def _controller_feedback():
    # Dobot CR V3: 1440-byte real-time feedback; no command is sent on this socket.
    import socket
    import struct
    host, port, *_ = robot.ConnectionParams()
    if int(port) != 29999:
        raise RuntimeError('当前连接不是已验证的Dobot CR反馈协议。')
    previous = None
    with socket.create_connection((host, 30004), timeout=3.0) as connection:
        deadline = time.monotonic() + 3.0
        for _ in range(2):
            packet = bytearray()
            while len(packet) < 1440:
                remaining = deadline - time.monotonic()
                if remaining <= 0:
                    raise RuntimeError('实机反馈读取超时。')
                connection.settimeout(remaining)
                part = connection.recv(1440 - len(packet))
                if not part:
                    raise RuntimeError('实机反馈连接已关闭。')
                packet.extend(part)
            length = struct.unpack_from('<Q', packet, 0)[0]
            marker = struct.unpack_from('<Q', packet, 48)[0]
            stamp = struct.unpack_from('<Q', packet, 32)[0]
            if length != 1440 or marker != 0x123456789ABCDEF:
                raise RuntimeError('实机反馈帧格式不匹配。')
            if previous is not None and stamp <= previous:
                raise RuntimeError('实机反馈时间戳未更新。')
            previous = stamp
        q = list(struct.unpack_from('<6d', packet, 192))   # ★真实关节角（v10定位，示教器交叉证实）；旧版误读432="连接基准+指令累加"的假值
        velocity = list(struct.unpack_from('<6d', packet, 480))
        mode = struct.unpack_from('<Q', packet, 24)[0]
        if not all(math.isfinite(v) for v in q + velocity):
            raise RuntimeError('实机反馈包含无效关节数值。')
        return q, velocity, mode


def _live_joints():
    if RDK.RunMode() != RUNMODE_RUN_ROBOT:
        raise RuntimeError('当前不是实机执行模式。')
    status, msg = robot.ConnectedState()
    if status != ROBOTCOM_READY:
        raise RuntimeError('机器人未就绪或已断连：' + str(msg))
    q, velocity, mode = _controller_feedback()
    # 阈值由 0.1 放宽到 1.0：实测静止时 J4/J3 的速度估计噪声可达 0.31°/s
    # （六轴角度 8 次采样完全相同），0.1 会把"其实已静止"误判为运动中而中止任务。
    if mode != 5 or max(abs(v) for v in velocity) > 1.0:
        raise RuntimeError('实机未处于使能静止状态，模式=%s。' % mode)
    return q


def _require_joints(expected):
    actual = _live_joints()
    if max(abs(a-b) for a,b in zip(actual, expected)) > 0.5:
        raise RuntimeError('关节反馈与预检状态不一致，停止后续命令。')


def _retreat_orientation_records(records):
    """加工点变姿态前退到 y=-750，变姿态后返回 y=-775。"""
    result = []
    previous = None
    for index, record in enumerate(records, 1):
        current = dict(record, values=record['values'][:])
        current['label'] = f'P{index}'
        if previous and previous['type'] == current['type'] == 'TCP':
            old, new = previous['values'], current['values']
            changed = pose_angle(invH(fanuc_values_to_pose(*old)) * fanuc_values_to_pose(*new)) > math.radians(.01)
            old_work, new_work = abs(old[1] + 775) < .001, abs(new[1] + 775) < .001
            if changed and (old_work or new_work):
                anchor = old if old_work else new
                retreat = dict(type='TCP', values=[anchor[0], -750., anchor[2]] + old[3:], singular=False,
                               label=f'P{index}前退让', require_linear=old_work)
                result.append(retreat)
                turn = dict(current, values=retreat['values'][:3] + new[3:], label=f'P{index}退让位换向')
                result.append(turn)
                current['singular'] = False
                current['require_linear'] = new_work
        result.append(current)
        previous = record
    return result


def _prepare_real_plan(records, start, deviation, single_method=None):
    RDK.setRunMode(RUNMODE_SIMULATE)
    try:
        RDK.Command('Trace', 'Off')
        robot.setJoints(start)
        if single_method is None:
            return _plan_continuous_trajectory(records, deviation, log)
        _enable_obstacle_checks()
        if robot.MoveJ_Test(start, start, minstep_deg=1) != 0:
            raise ValueError('起始姿态碰撞：' + _collision_details())
        values = records[0]['values']
        method, fallback = single_method, False
        if method not in ('MoveJ','MoveL'):
            raise ValueError('未知单点运动类型。')
        end = None
        waypoints = []
        if method == 'MoveL':
            end, _ = _linear_path_endpoint(start, fanuc_to_pose(*values))
            if end is not None:
                # v13：单点 MoveL 同样不信任驱动 MOVL（纯J6自转也一样，关节插值=同一路径），
                # 改细分途经点+MoveJ 执行
                waypoints = _linear_waypoints(start, fanuc_to_pose(*values))
                if waypoints:
                    log('单点 MoveL 改细分执行：%d 个途经点（步长≤%.0fmm）。' % (len(waypoints), LINEAR_SUBSTEP_MM))
                    log('单点 MoveL 途经跳（共%d跳）：%s' % (len(waypoints), [[float('%.2f' % v) for v in w] for w in waypoints]))
        if end is None:
            end = _obstacle_joint_target(start, values, deviation if method=='MoveL' else None)
            fallback, method = method=='MoveL', 'MoveJ'
        plan = [dict(method=method,joints=end,special=False,fallback=fallback,rewinds=[],j6_delta=None,waypoints=waypoints)]
        _verify_obstacle_plan(start, plan)
        return plan
    finally:
        robot.setJoints(start)
        RDK.Render(True)
        RDK.setRunMode(RUNMODE_RUN_ROBOT)  # 旧版 L615 有此行：预检后必须切回实机模式，否则 _live_joints 直接拒执行


def _wait_controller_static(max_wait_s=20.0, vel_threshold=0.5, samples=5, interval=0.3):
    """轮询30004反馈直到六轴静止（连续samples次速度<阈值），返回(关节, 是否静止)。

    v14o：断连分支以 samples=3/interval=0.2 调用（短跳≈1s，5×0.3s 静止确认占每跳
    尾部 ~1.5s，是停顿税大头）；默认 5×0.3s 供正常路径；20s 静止上限（真断连护栏）不动。"""
    t0 = time.time()
    quiet = 0
    last = None
    while time.time() - t0 < max_wait_s:
        actual, velocity, _mode = _controller_feedback()
        last = actual
        if max(abs(v) for v in velocity) < vel_threshold:
            quiet += 1
            if quiet >= samples:
                return last, True
        else:
            quiet = 0
        time.sleep(interval)
    return last, False


def _wait_arrival_then_static(target_joints, max_wait_s=20.0):
    """v14u：目标锚定的到位等待——直发后不再猜「起步了没」，只等「到没到」。

    背景（v14t 10:38 P9 实测）：直发指令起步延迟可 >6s，让位 6s 耗尽判「未执行」
    停止后，指令仍被控制器自行执行到精确目标（善后实测 J2 +10°/J3 +20°，余轴不动，
    宏未重发）——「起点静止」与「完成静止」在反馈上不可区分，位置对目标才是唯一
    可靠锚点（速度判据出局：三场停时 J4 0.06~0.42°/s 均为低于阈值的保持抖动）。
    本函数：距目标关节 ≤MOVL_ARRIVE_TOL_DEG 且速度<0.5°/s → 到位完成（此时已在
    目标，无需再做常规静止确认）；每 5s 一行进度日志（顺带实测真实延迟）；
    上限 MOVL_ARRIVE_WAIT_S 超时报「疑似未执行」停待判读；不重发铁律不变。
    target_joints=None → 退化为 _wait_controller_static()，行为与原先完全一致。"""
    if target_joints is not None:
        t0 = time.time()
        t_note = t0
        while True:
            fb = _controller_feedback()
            err = max(abs(a - b) for a, b in zip(fb[0], target_joints))
            if err <= MOVL_ARRIVE_TOL_DEG and max(abs(v) for v in fb[1]) < 0.5:
                log('MovL 直发到位确认：距目标关节%.2f°（%.1fs），验收继续。'
                    % (err, time.time() - t0))
                return fb[0], True
            if time.time() - t0 >= MOVL_ARRIVE_WAIT_S:
                raise RuntimeError(
                    'MovL 直发%.0fs仍未到位（距目标关节%.2f°），疑似未执行，停止待判读。'
                    % (MOVL_ARRIVE_WAIT_S, err))
            if time.time() - t_note >= 5.0:
                log('MovL 直发等待到位：%.0fs，距目标关节%.2f°，续等（不重发，上限%.0fs）。'
                    % (time.time() - t0, err, MOVL_ARRIVE_WAIT_S))
                t_note = time.time()
            time.sleep(0.5)
    return _wait_controller_static(max_wait_s=max_wait_s)


MOVE_OFFSET_TOL = 0.5   # 闭环补偿后的到位容差（°）


TCP_TOOL_NAME = 'CR5_TCP_126mm'
FLANGE_TOOL_NAME = '_CR5_FLANGE_DIRECT_TEMP'
_tool_window_depth = 0


def _same_tool_pose(a, b):
    return max(abs(a[r, c] - b[r, c]) for r in range(4) for c in range(4)) < 1e-7


def _named_tool(name, pose):
    matches = [it for it in robot.Childs()
               if it.Type() == ITEM_TYPE_TOOL and it.Name() == name]
    if len(matches) > 1:
        raise RuntimeError('重复 TCP 工具条目：' + name)
    if matches:
        tool = matches[0]
        if not _same_tool_pose(tool.PoseTool(), pose):
            raise RuntimeError('TCP 工具定义不符，停止待核对：' + name)
        return tool
    return robot.AddTool(pose, name)


def _restore_tool(pose, linked_tool=None):
    """Restore the original item link when possible, and never swallow failure."""
    for attempt in range(2):
        try:
            robot.setPoseTool(linked_tool if linked_tool is not None and linked_tool.Valid() else pose)
            if not _same_tool_pose(robot.PoseTool(), pose):
                raise RuntimeError('PoseTool 恢复后读回不一致')
            return
        except Exception as exc:
            if attempt == 1:
                raise RuntimeError('工具恢复失败，禁止继续运动：' + str(exc)) from exc


def _single_move_settle(method, target, require_joints=True, expect_target=None, flange_space=False, _retry=0):
    """发指令并确认到位——v14w39 窗口版入口：flange_space 时单位变换+藏把手覆盖
    【整个 settle 生命周期】（发送+断连恢复+到位等待）。旧版只包 RPC 一次调用：假断连
    抛出时窗口即关、把手提前回来，RoboDK 本地退化动画在弧 66% 被碰撞检测掐停→模型冻在
    撞点、红显常驻→收口 MoveJ 被拦死（10-22 四次实录含 v14w38）。"""
    global _tool_window_depth
    if not flange_space or _tool_window_depth:
        # A controlled retry already runs inside the outer tool window.
        # Only the outer owner may restore the original TCP.
        return _settle_core(method, target, require_joints, expect_target, flange_space, _retry)
    _ensure_canonical_tool()
    _win_tp = robot.PoseTool()
    _win_link = robot.getLink(ITEM_TYPE_TOOL)
    _win_handle = RDK.Item('门把手_bs1')
    _win_visible = _win_handle.Visible() if _win_handle.Valid() else None
    _flange_tool = _named_tool(FLANGE_TOOL_NAME, eye(4))
    _tool_window_depth += 1
    try:
        robot.setPoseTool(_flange_tool)
        if not _same_tool_pose(robot.PoseTool(), eye(4)):
            raise RuntimeError('法兰工具切换失败，未发送运动指令')
        if _win_visible is not None:
            _win_handle.setVisible(False)
        return _settle_core(method, target, require_joints, expect_target, True, _retry)
    finally:
        try:
            _restore_tool(_win_tp, _win_link)
        finally:
            _tool_window_depth -= 1
            if _win_visible is not None:
                _win_handle.setVisible(_win_visible)


def _settle_core(method, target, require_joints, expect_target, flange_space=False, _retry=0):
    """发一条运动指令并确认到位（v10：反馈字段已校正）。

    v14r：require_joints=False 仅供 MovL 直发调用点使用——断连分支的关节级 0.5°
    校验让位给外层法兰级粗验收（≤8mm/≤1°）+MoveJ 微纠偏收口（v14q 09:57 实机
    教训：MovL 直发必触发假断连，0.95° 固有残差在断连分支内即被拦停，外层验收
    根本没执行到）。其余护栏不变：20s 静止上限、重连失败仍停。

    v14u：断连分支改目标锚定到位等待 _wait_arrival_then_static——上限 60s 每 5s
    进度日志；超时报「疑似未执行」停。不重发铁律不变。

    v14w37：直发=【法兰位姿传递 + flange_space 单位变换窗口】双件套——
    ①传位姿（调用方 invH(PoseFrame)*SolveFK(净化关节) 自算）：MoveL 的动画按位姿空间
    直线走=认证路径，根治旧 MoveL(关节) 的关节弧动画扫进圆柱假碰撞冻死（10-22 两次实录）；
    ②发送 RPC 窗口内 PoseTool 置单位变换：MoveL(位姿) 的可达校验/语义都按 TCP 空间做，
    不切工具则法兰位姿被当 TCP 反推（P8 反推法兰 z=744 爆臂展 ⇒ TargetReachError，
    10-22 11:18 实录）；单位变换下校验空间=法兰空间，数字逐位=金标准（实证 0 偏差）。
    动画窗口内直线途经点 12/12 无碰撞（单位变换工具下实测）。
    v14w38：窗口内追加隐藏把手——驱动断连瞬间 RoboDK 本地退化关节动画（会撞圆柱的
    那条弧）是三次冻结的真凶；藏把手=对假路径的检测放行（实测弧中点/冻结姿态
    显隐 True/False 翻转），真直线 1mm 检查本来就 0 碰撞。

    v14w20：受控补发（一次性）——驱动连接恰死在发送时刻时 SendJointMovJ 会静默
    丢弃不发送（反汇编：CONNECTED=False 直接 return False；2026-10-15 09:51 P25
    实发：断连后臂停在发送前位置、误差127.8°）。补发条件（全部满足才补，且全程
    至多一次）：①失败 ②30004 独立反馈证明【零位移】（仍在发送前关节 ≤0.5°）
    ③ensure_connected() 重连成功。指令已上线/延迟执行/落点异常的场景均不满足
    ②（有位移）不会触发——保留原「不重发」语义。历史上"晚执行"案例（v14t）
    后经控制器日志证实为面板拖动误判，非队列延迟。

    历史结论：驱动一直正确执行绝对关节目标；真实关节角在偏移192。"""
    try:
        _start_q = None
        try:
            _start_q = _controller_feedback()[0]
        except Exception:
            _start_q = None
        getattr(robot, method)(target)   # v14w39：flange 窗口已上移至 _single_move_settle 包装层
    except StoppedError as exc:
        if str(exc).strip() != 'Robot not connected':
            raise
        # v14o 静默重连：假断连是本环境常态（每条 MoveJ 指令结束后都可能误报）；30004
        # 反馈通道独立于驱动连接，静止确认与重连并行进行，压缩跳间停顿税。
        # 护栏不变：未自然收尾（20s 上限）仍停、落点仍 0.5° 校验、重连失败仍停。
        log('驱动报断连——等待收尾与后台重连并行进行…')
        import threading as _st
        reconnected = []
        def _bg_reconnect():
            for _r in range(3):
                if ensure_connected():
                    reconnected.append(True)
                    return
                time.sleep(1.0)
        _rt = _st.Thread(target=_bg_reconnect, daemon=True, name='silent_reconnect')
        _rt.start()
        # v14u：到位等待下沉在断连分支（MovL 直发永远走本分支——v14s 教训）——
        # 目标锚定：距目标≤2°且静止=完成，不猜起步。非 MovL 直发退化为常规静止确认。
        try:
            actual, is_static = _wait_arrival_then_static(expect_target)
        except RuntimeError as _arr_exc:
            # v14w20：直发「疑似未执行」——零位移+重连成功 ⇒ 补发一次（指令未上线实证）
            if (_retry < 1 and _start_q is not None
                    and max(abs(a - b) for a, b in zip(_controller_feedback()[0], _start_q)) <= MOVE_OFFSET_TOL
                    and ensure_connected()):
                log('直发疑似未执行且零位移（仍在起点）——判定指令未上线，补发一次（v14w20）。')
                return _single_move_settle(method, target, require_joints, expect_target,
                                           flange_space, _retry=_retry + 1)
            raise
        if not is_static:
            raise RuntimeError('驱动报断连后等待%.0fs仍未静止，停止。' % 20.0) from exc
        if require_joints:
            err = max(abs(a - b) for a, b in zip(actual, target))
            if err > MOVE_OFFSET_TOL:
                # v14w20：MoveJ 类「断连收尾后未到位」——零位移+重连成功 ⇒ 补发一次
                if (_retry < 1 and _start_q is not None
                        and max(abs(a - b) for a, b in zip(actual, _start_q)) <= MOVE_OFFSET_TOL
                        and ensure_connected()):
                    log('断连后零位移（仍在起点）——判定指令未上线，补发一次（v14w20）。')
                    return _single_move_settle(method, target, require_joints, expect_target,
                                               flange_space, _retry=_retry + 1)
                raise RuntimeError('断连收尾后未到位：目标%s，实测%s（误差%.2f°），停止待判读。'
                                   % (['%.2f' % v for v in target], ['%.2f' % v for v in actual], err)) from exc
        _rt.join(timeout=4.0)
        if not reconnected:
            raise RuntimeError('已到位但驱动重连失败，停止后续指令。') from exc
        log('驱动断连但运动已自然完成到位；已重连驱动，继续。')
        return
    actual, is_static = _wait_controller_static()
    if not is_static:
        raise RuntimeError('指令返回后等待静止超时（20s），停止。')
    if require_joints:
        err = max(abs(a - b) for a, b in zip(actual, target))
        if err > MOVE_OFFSET_TOL:
            raise RuntimeError('落点偏差%.2f°：目标%s，实测%s，停止待判读。'
                               % (err, ['%.2f' % v for v in target], ['%.2f' % v for v in actual]))
    return


MOVE_OFFSET_TOL = 0.5   # 到位容差（°）：反馈字段校正后，超过即停止待判读


# v13（方案B）：驱动 MOVL 执行层已判死（3 次实机断连指纹 + .pyc 反汇编直连无收尾），
# 所有 MoveL 执行全部替换为「细分途经点 + MoveJ」。作业面短段（≤ TRANSIT_DIRECT_MAX_MM）
# 用 MoveL 指令的 1mm 逆解采样出 ≤ LINEAR_SUBSTEP_MM 的途经关节序列，MoveJ 逐跳执行；
# 过渡段长段优先 MoveJ 直达（须过 TCP 偏离≤max_deviation 且整弧 MoveJ_Test 碰撞检查），
# 不满足才退回细分。预检层 MoveL_Test@1mm 保留：仍是「这一段能不能走直线」的权威筛选器。
TRANSIT_DIRECT_MAX_MM = 300.0   # 超过此段长的 TCP 段视为自由空间过渡段，尝试 MoveJ 直达
LINEAR_SUBSTEP_MM = 20.0        # 作业面细分步长：v14m(40mm) 实机碰撞实证弦误差可吃掉真裕度（轴线距199.9-半径180≈19.9mm），回 20mm 安全基准（v14k 两度全通过）；途经点弦误差 <0.5mm

MOVL_DIRECT_MAX_MM = 210.0   # v14w35（10-22）：150→210——150 是 v14p 照当时谱系（最长≈120mm）取的设计余量，非事故判死值；210 覆盖 200mm 工艺段一指令（y=-719 线翻转点→x=-100），留 FP 边界余量。路径背书不变（认证直线+整段复核）；更长直线段仍走细分
# ★★★ v14w（2026-10-13 16:08）：【禁直发名单清空 = 恢复 P9 直发】+ 发送位姿数字净化。
#   v14v4 按点号拦 P9 是在 -30001 真凶查明前的临时措施（且拦下分支会落空——随名单清空，
#   该落空分支变为不可达死码，留档不删）。真凶 = 控制器 MovL 参数校验拒收【参数形态】
#   （-0.000000 / +90.000000 / -0.000000，见 LOG_VERSION 处实录），不是几何、不是段长：
#   同目标 15:55:51 单步直发实证 return 0、1.1s 到位。净化失败 ⇒ 本段自动改走细分（安全回落）。
# 想再拦某点：改回 (9,) 即可（注意拦下分支的落空缺陷仍在，见 P2P_LESSONS.md）。
MOVL_DIRECT_BLOCK_POINTS = ()
MOVL_FLANGE_TOL_MM = 8.0     # v14q 直发 MovL 法兰位置粗验收容差：控制器 MovL 固有落点残差实测 4.61mm（v14p 首航）/5.5mm（v14l）双样本，取实测+裕量；超此值=落点异常真停
MOVL_FLANGE_TOL_DEG = 1.0    # v14q 直发 MovL 法兰姿态粗验收容差（实测 0.616°+裕量）；通过后 MoveJ 微纠偏收口到关节级 0.5° 内
MOVL_ARRIVE_WAIT_S = 60.0    # v14u MovL 直发到位等待上限：目标锚定（距目标≤2°且静止即完成），不猜起步——v14t 10:38 实测 P9 起步延迟>6s、指令事后自行执行完；60s 为 10 倍裕量，每5s进度日志实测真实延迟，超时按未执行停待判读
MOVL_ARRIVE_TOL_DEG = 5.0    # v14u 到位判定关节距离阈（°）；v14w30 2→5：tool=182 构型下 ~5mm 固有误差映射关节达 2.58°（10-21 P8 实证），阈外即误判未执行——粗验收前哨放宽，法兰级粗验收(≤8mm/≤1°)+MoveJ收口紧随其后罩终点；此处不走 MOVE_OFFSET_TOL=0.5°（require_joints=False 路径，护栏语义不降级）

# v14w22：实机关节限位（与 RoboDK 模型 ±360 取交集）。依据：J1=193.59 两次被控制器
# -40001 拒收（10-15 P25）；J6=190.84 return 0 ✓；J5=177.6 实机走成 ✓（故 J5=180 非
# 某些资料的 ±120）；J3 取模型更紧的 ±160。规划期过滤，保证预检路径=实发路径。
# v14w23：J4 190→150——J4=-189.70 被控制器 -40004（自干涉 PoseSelfInterference）拒收；
# -168 族中途自干涉保护停机；实证安全族 |J4|≤95，150 留 55° 余量。
REAL_JOINT_LIMITS = (180.0, 180.0, 160.0, 150.0, 180.0, 360.0)

# v14w26：实机自干涉组合区（控制器 PoseSelfInterference 的 J4×J5 耦合，-40006）。
# 实录：|J4|=115.5×|J5|=173.1 与 |J4|=109.4×|J5|=171.5 均拒；|J4|=83.2×|J5|=177.6 通过。
# 阈值取中：|J4|>100 且 |J5|>165 视为禁区（两端各留 ~9°/~8° 实证余量）。
REAL_INTERFERE_J4_MAX = 100.0
REAL_INTERFERE_J5_MIN = 165.0


def _real_interfere_combo(q):
    """v14w26：关节是否落入实机自干涉组合禁区（J4×J5 耦合，控制器 -40006）。"""
    return abs(q[3]) > REAL_INTERFERE_J4_MAX and abs(q[4]) > REAL_INTERFERE_J5_MIN


def _real_limit_ok(q, lower, upper):
    """v14w22：关节目标是否同时满足模型限位与实机限位。"""
    for j in range(min(6, len(q))):
        lo = max(float(lower[j]), -REAL_JOINT_LIMITS[j])
        hi = min(float(upper[j]), REAL_JOINT_LIMITS[j])
        if not lo <= float(q[j]) <= hi:
            return False
    return True


def _movl_digit_safe_joints(q_target):
    """v14w：直发位姿数字净化 —— 控制器 MovL 参数校验 -30001 防御。

    实证（控制器 logs/all/log）：
      11:38:20 拒收 MovL(-0.000000,…,300.000000,90.000000,0.000000,-0.000000)
               → [MovL#820] the type of params is wrong: -30001
      15:55:51 接受 MovL(0.000000,…,299.999986,89.999995,-0.000003,0.000000) → return 0
    触发器（同目标、不同关节末位 ⇒ 不同参数形态 ⇒ 校验翻转）：
      x 负零/极小负 · rx 恰=+90.000000 · **三角(rx/ry/rz)负零——ry=-0 是 -30005 实锤**
      （10-15 09:16 与 10-14 拒收样本共同点；接受样本 ry 均为 +0）· rz=+180（保留防御）
      —— 同时设防，且只在零/边界区动手：
      · x ∈ (-0.01, 0.001) mm → 推到 ≥ +0.001（FK 位置与欧拉约定无关，可靠）
      · rx ∈ [89.999, 90.001] → 拉出该区（Pose_2_Fanuc 的 rx 与两份实录一致）
      · rz 为负零 (-0.0) → 推离
    手法：对发送关节贪心微扰（步长 0.0005°→0.05°，单关节累计 ≤0.05°，末端位移 ≲0.6mm
    ≪ 圆柱真裕度 19.9mm ≪ 法兰验收 8mm）；到位/法兰验收/MoveJ 收口仍对【原始认证关节】
    判定，收口回认证构型 —— 几何语义不变。P5 类非边界参数零扰动（首查即过，原样返回）。
    返回 (send_q, note)：无违规=(原关节,None)；成功=(微扰关节,说明)；失败=(None,原因)。"""
    def _digits(q):
        # v14w19：先按驱动下发格式（6位小数）定型再判——控制器校验的是字符串形态；
        # 客户端 Fanuc 与驱动在零点附近的正负号约定不一致，故三角一律推离零域。
        # v14w24：净化微扰可能把限位边界关节（如 J6=-360.00）推出模型限位，
        # SolveFK 会抛 TargetReachError——捕获后返回 None=不可行候选（评分置顶永不选中）。
        try:
            return [float('%.6f' % v) for v in Pose_2_Fanuc(robot.SolveFK(q))]
        except Exception:
            return None

    def _score(vals):
        if vals is None:
            return 1e9   # 越界候选：永不优于当前
        x, rx, ry, rz = vals[0], vals[3], vals[4], vals[5]
        s = 0.0
        if -0.01 < x < 0.001:                      # 零附近（含 -0.000000）且未达 +0.001
            s += (0.001 - x) / 0.001
        if 89.999 <= rx <= 90.001:                 # 恰卡 +90 边界（含 90.000000 整）
            s += (rx - 89.999) / 0.001
        # v14w19：三角必须整体离开零域 ≥0.001°——"-0.000000"形态是 -30005 实锤
        #（10-15 09:16/09:35 两次实录 ry 打印 -0.000000 均拒；-2e-7 打印即 -0.000000
        #  而浮点 !=0.0 会漏判；推离零域后客户端/驱动符号一致为正）
        for v in (rx, ry, rz):
            if abs(v) < 0.001:
                s += 1.0 + (0.001 - abs(v)) / 0.001
        if rz >= 179.999:                          # rz=+180 疑似越界（保留防御）
            s += 1.0 + (rz - 179.999) / 0.001
        return s

    base = list(q_target)
    cur = _score(_digits(base))
    if cur <= 0.0:
        return q_target, None
    q = list(base)
    solved = False
    for step in (0.0005, 0.002, 0.01, 0.05):
        improved = True
        while cur > 0.0 and improved:
            improved = False
            for j in range(6):
                for sgn in (1.0, -1.0):
                    q2 = q[:]
                    q2[j] += sgn * step
                    if abs(q2[j] - base[j]) > 0.05 + 1e-9:
                        continue
                    sc = _score(_digits(q2))
                    if sc < cur - 1e-12:
                        q, cur, improved = q2, sc, True
                        break
                if improved:
                    break
        if cur <= 0.0:
            solved = True
            break
    if not solved:
        return None, '发送位姿净化失败（边界参数 x/rx/rz 微调不出安全区）'
    touched = ['%s%+.4f' % ('J%d' % (k + 1), q[k] - base[k]) for k in range(6)
               if abs(q[k] - base[k]) > 1e-9]
    return q, '发送关节微扰 %s°（Δmax 对应末端 ≪1mm）：规避 -30001 边界参数；验收/收口仍回认证构型' \
        % ' '.join(touched)


def _movl_flange_accept(joints_now, joints_target):
    """v14q：直发 MovL 落点的法兰位姿级粗验收。

    v14p 首航实证：控制器 MovL 固有落点残差 ~5mm/0.6° 级（v14p 4.61mm/0.616°、v14l 5.5mm，
    双样本跨版本一致）——关节级 0.5° 判据会把正常落点误判为事故。改用法兰语义验收：
    FK(实测) vs FK(目标)，位置≤MOVL_FLANGE_TOL_MM 且姿态≤MOVL_FLANGE_TOL_DEG 即过；
    过后在 _execute_checked_real 里发一条 MoveJ 微纠偏收口（关节级 0.5° 校验罩住终点）。
    超容差=落点异常（构型翻转/卡住/送错目标），照旧抛 RuntimeError 即停待判读。"""
    _f_now = invH(robot.PoseFrame()) * robot.SolveFK(joints_now)      # 法兰位姿（无工具）
    _f_tgt = invH(robot.PoseFrame()) * robot.SolveFK(joints_target)
    _d = _f_now * invH(_f_tgt)
    _mm = norm(_d.Pos())
    _deg = math.degrees(pose_angle(_d))
    return _mm, _deg


def _movl_direct_ready():
    """v14p 法兰补偿MOVL 开关是否可用：GUI 变量已建（正常运行）才开；
    离线 verify 的 exec 命名空间里没有 real_movldirect_var（NameError），
    自动回 False——离线验证的计划/指纹与该开关无关（规划层零改动）。"""
    try:
        return isinstance(real_movldirect_var, tk.BooleanVar)
    except Exception:
        return False


MOVE_SEGMENT_MAX_DEG = 64.0  # 每瓣最大关节跨度：驱动约8秒无完成回报即断连，20°/s下64°≈3秒，留足裕量


J6_SPIN_SEGMENT_DEG = 60.0   # MoveL 纯J6自转段分瓣跨度（无平移时关节插值=笛卡尔路径）


def _is_pure_j6_spin(start, target):
    """MoveL 目标仅 J6 变化（J1~J5 不动）：关节插值与笛卡尔路径重合，可精确分瓣。"""
    return max(abs(a - b) for a, b in zip(start[:5], target[:5])) < 1e-6


def _move_with_completion_check(method, target, allow_split=True):
    """长运动分瓣执行（v9）：驱动对单条指令约8秒无完成回报就断连（本环境常态，
    test.py 同款假报，它每段部在几秒内完成所以从没撞上）；大跨度关节运动沿
    预检验证过的同一条关节直线剖成若干瓣，每瓣都在死线内完成，路径不变，
    仅增设停顿点。MoveL 纯J6自转段同理分瓣；带平移 MoveL 与小跨度段保持原样。"""
    if not allow_split:
        # v11: 单点运动/关节运动不分瓣，恢复一指令直达（到位校验与假断连容忍保留）
        _single_move_settle(method, target)
        return
    try:
        start = _live_joints()
        total = max(abs(float(b) - float(a)) for a, b in zip(start, target))
    except Exception:
        start, total = None, None
    if method == 'MoveJ' and total is not None and total > MOVE_SEGMENT_MAX_DEG:
        pieces = int(math.ceil(total / MOVE_SEGMENT_MAX_DEG))
        log('长运动分瓣：跨度%.1f° → %d 瓣执行（同一关节直线，仅增设停顿点）。' % (total, pieces))
        for k in range(1, pieces + 1):
            way = [a + (b - a) * k / pieces for a, b in zip(start, target)]
            _single_move_settle('MoveJ', way)
            _require_joints(way)  # 瓣间校验到位，也给驱动链路留出响应时间
        return
    if (method == 'MoveL' and total is not None and _is_pure_j6_spin(start, target)
            and total > J6_SPIN_SEGMENT_DEG):
        pieces = int(math.ceil(total / J6_SPIN_SEGMENT_DEG))
        log('J6自转分段：跨度%.1f° → %d 段MoveL（纯自转，路径与笛卡尔路径重合）。' % (total, pieces))
        for k in range(1, pieces + 1):
            way = [a + (b - a) * k / pieces for a, b in zip(start, target)]
            _single_move_settle('MoveL', way)
            _require_joints(way)
        return
    _single_move_settle(method, target)


_real_running = False  # 2026-10-09 补回：旧版 L510 有此初始化，升级版漏带导致点击即 NameError 静默炸裂


def _ensure_canonical_tool():
    """v14w17：工具坐标守护——检测到 identity(0)（存档僵尸/直发残留）自动恢复规范值并大声记日志。
    实发两次：2026-10-14 18:2x、2026-10-15 09:0x（归零→种子/P2 预检异常、P5 直发异常）。
    v14w39：同时恢复被直发窗口残留隐藏的门把手（GUI 中途被杀会留下隐藏态→预检漏检）。
    每次执行入口 + 程序启动各调一次；非零值不干预（可能正在被人工调整）。"""
    if _tool_window_depth:
        return False  # Do not undo the intentional identity TCP during MOVL.
    pose = robot.PoseTool()
    fixed = False
    canonical = Fanuc_2_Pose(list(CANONICAL_TOOL))
    if _same_tool_pose(pose, eye(4)) or _same_tool_pose(pose, canonical):
        tcp = _named_tool(TCP_TOOL_NAME, canonical)
        _restore_tool(canonical, tcp)
    if _same_tool_pose(pose, eye(4)):
        log('⚠️ 工具坐标为0（存档残留/直发残留）——已自动恢复 [0,0,126]，请确认后再跑。')
        fixed = True
    try:
        _gh = RDK.Item('门把手_bs1')
        if _gh.Valid() and not _gh.Visible():
            _gh.setVisible(True)
            log('⚠️ 门把手网格处于隐藏态（直发窗口残留）——已恢复显示。')
            fixed = True
    except Exception:
        pass
    return fixed


def _execute_checked_real(data, single_method=None):
    global _real_running
    log('【入口】_execute_checked_real：%d 点，single_method=%s' % (len(data) if data is not None else -1, single_method))
    if _real_running:
        log('已有实机任务正在执行。')
        return
    _real_running = True
    completed = 0
    movl_direct = False  # v14p：入口预置，防异常早于赋值时 except 块二次 NameError（v14l 教训）
    try:
        _ensure_canonical_tool()  # Failure must pass through task cleanup.
        log('开始校验录入数据…')
        records = _validated_records(data)
        log('录入数据校验通过：%d 点。' % len(records))
        if single_method is None and len(records) > 1:
            expanded = _retreat_orientation_records(records)
            log('连续轨迹：%d个录入点展开为%d个执行点（含姿态退让）。' % (len(records), len(expanded)))
            records = expanded
        deviation = float(real_deviation_var.get())
        if not math.isfinite(deviation) or deviation < 0:
            raise ValueError('允许偏离必须为非负有限数。')
        log('偏离上限 %.1f mm，检查机器人连接…' % deviation)
        if not ensure_connected():
            return
        start = _live_joints()
        log('实机当前关节：%s' % ['%.2f' % v for v in start])
        # 长预检/运动期间 RoboDK 主程序忙或不消费驱动输出，驱动链路会饿死断开（15:20:56 P1 中途断连同因）。
        # 保活线程用独立 API 连接（避免被 MoveJ 阻塞主连接），每2秒一次 ConnectedState（只读），
        # 贯穿预检+执行全程，直到任务结束才停（v7 错在预检后就停，P1 运动中饿死驱动）。
        import threading as _th
        _keepalive_stop = _th.Event()
        def _driver_keepalive():
            n = 0
            _ka_rdk = Robolink()
            _ka_robot = _ka_rdk.Item('', ITEM_TYPE_ROBOT)
            while not _keepalive_stop.wait(2.0):
                n += 1
                try:
                    s, _m = _ka_robot.ConnectedState()
                    if s < 0:
                        log('【保活】第%d次发现驱动掉线（%s），已请求重连。' % (n, _m))
                        _ka_robot.Connect()
                except Exception:
                    pass  # 主程序忙时 API 调用可能慢/超时，下一轮再试
        _ka_thread = _th.Thread(target=_driver_keepalive, daemon=True, name='driver_keepalive')
        _ka_thread.start()
        log('已启驱动保活（贯穿预检+执行）。')
        frame, tool = robot.PoseFrame(), robot.PoseTool()
        log('开始台子/地面避障预检，尚未发送运动指令。')
        plan = _prepare_real_plan(records, start, deviation, single_method)
        # 保活线程不在此处停：执行阶段同样需要（v7 教训）
        # 预检后复核：驱动必须就绪且关节与预检起始一致，否则取消。
        if not ensure_connected():
            log('预检后驱动断连，重连未成功，取消执行。')
            return
        _require_joints(start)
        log('预检后连接复核通过，准备发运动指令。')
        # v14w22：实机限位最后防线（规划器已过滤，此处兜底拦截任何漏网目标）
        _lo, _hi, _ = robot.JointLimits()
        _lo, _hi = _lo.list(), _hi.list()
        for _i, _step in enumerate(plan, 1):
            if not _real_limit_ok(_step['joints'], _lo, _hi):
                raise ValueError('段%d 目标关节超出实机限位：%s（规划期应已过滤，此为最后防线）'
                                 % (_i, ['%.2f' % v for v in _step['joints']]))
        for before, after in ((frame, robot.PoseFrame()), (tool, robot.PoseTool())):
            error = invH(before)*after
            if norm(error.Pos()) > 0.01 or pose_angle(error) > math.radians(0.01):
                raise RuntimeError('预检期间工具或参考坐标系改变，取消执行。')
        robot.setSpeed(ROBOT_SPEED)
        RDK.Command('Trace','Reset')
        RDK.Command('Trace','On')
        expected = start
        # v14k：停用长运动分瓣（split_moves 恒 False）。2026-10-12 实测日志坐实：假断连与跨度无关，
        # 60°/95°/169°/180° 的瓣与 20mm 途经点每条指令都在断，分瓣已不防任何东西，只剩每瓣一轮
        # 等待+重连停顿税；_single_move_settle 断连容忍（_wait_controller_static 20s 静止上限）
        # 罩得住单条长指令的收尾（20°/s 下 180°≈9s<20s）。分瓣机制与常量原样留档，遇真断连指纹
        # （未自然收尾/未到位）随时把本行改回 single_method is None and len(records) > 1 即可恢复。
        split_moves = False
        movl_direct = bool(real_movldirect_var.get()) if _movl_direct_ready() else False
        if movl_direct:
            log('【v14w41】法兰补偿MOVL默认开启：短直线段（≤%.0fmm、姿态恒定≤0.5°）一指令直发驱动 MOVL（工具补偿；发送关节自动净化规避控制器 -30001/-30005 边界参数；落点法兰级粗验收≤%.0fmm/%.1f°+MoveJ微纠偏收口+到位等待≤%.0fs 目标锚定·关节阈5°；J6±360边界换同角表示；同位姿换姿优先MoveJ分支直达；规划与预检不变；净化失败自动改走细分；断连零位移时受控补发一次；关节目标实机限位(180/180/160/150/180/360)规划期过滤；J4×J5 自干涉组合区(-40006)规划期禁选；工具=126mm）。'
                '★ 禁直发名单=%s（空=全部可直发；净化失败的点自动回落细分）。' % (MOVL_DIRECT_MAX_MM, MOVL_FLANGE_TOL_MM, MOVL_FLANGE_TOL_DEG, MOVL_ARRIVE_WAIT_S, MOVL_DIRECT_BLOCK_POINTS))
        for i, step in enumerate(plan, 1):
            for rewind in step['rewinds']:
                _require_joints(expected)
                _move_with_completion_check("MoveJ", rewind, split_moves)
                _require_joints(rewind)
                expected = rewind
            _require_joints(expected)
            waypoints = step.get('waypoints') or []
            if step['method'] == 'MoveL' and not waypoints:
                # 理论不可达：v13 起所有 MoveL 步都带细分途经点；不带则说明规划层契约被破坏
                raise RuntimeError(f"P{i}：MoveL 步缺少细分途经点，拒绝发送驱动 MOVL（已判死）。")
            seg_mm = seg_rot = None
            if movl_direct and step['method'] == 'MoveL' and waypoints:
                # 仅开关开启时才算（两次 FK 的 API 往返）；开关关/离线 verify 零开销
                _seg_rel = _trajectory_pose(step['joints']) * invH(_trajectory_pose(expected))
                seg_mm, seg_rot = norm(_seg_rel.Pos()), pose_angle(_seg_rel)
            direct_ready = (movl_direct and i not in MOVL_DIRECT_BLOCK_POINTS
                            and seg_mm is not None
                            and seg_mm <= MOVL_DIRECT_MAX_MM
                            and seg_rot <= math.radians(0.5))
            _send_q = step['joints']
            if direct_ready:
                # v14w：发送前数字净化——控制器 -30001 拒的是【参数形态】不是几何（LOG_VERSION
                # 处 11:38 拒收 / 15:55 接受两份实录）。净化只在零边界区微调发送关节；
                # 净化失败 ⇒ direct_ready=False ⇒ 落到 elif waypoints 走细分（安全回落）。
                _send_q, _purge_note = _movl_digit_safe_joints(step['joints'])
                if _send_q is None:
                    log('P%d：⛔ %s ⇒ 改走细分途经点路径。' % (i, _purge_note))
                    direct_ready = False
                elif _purge_note:
                    log('P%d：%s' % (i, _purge_note))
            if direct_ready:
                # v14p 法兰补偿MOVL：驱动 MOVL 无工具补偿、按法兰执行（v14l 11:30 实证停点法兰=
                # 命令TCP目标，差仅5.5mm）——将错就错：把本步构型的【法兰位姿】直接当笛卡尔目标
                # 发给控制器，法兰被精确送到位，物理工具尖端（182mm，v14w27 实测）随之落在认证
                # 直线上。姿态恒定段法兰线=TCP线平移常向量，扫掠包络与细分路径一致。
                # v14w36/37 演进：v14w36 只改传位姿（不切工具）⇒ MoveL(位姿) 按 TCP 空间
                # 校验，P8 法兰位姿被反推到 z=744 爆臂展 TargetReachError（11:18 实录）；
                # v14w37 = 位姿传递（动画=认证直线，根治关节弧假碰撞冻死）+ 发送窗口单位
                # 变换（校验/数字=法兰空间）；柜子实收参数与旧金标准逐位一致（0 偏差）。
                log(f"P{i}：v14w 法兰补偿MOVL：段长{seg_mm:.1f}mm（姿态变化{math.degrees(seg_rot):.2f}°），收起 {len(waypoints)} 个细分途经点，一指令直发（发法兰位姿=自算FK+单位变换窗口，发送关节已净化；v14w37）。")
                # v14r：require_joints=False——假断连分支的关节级 0.5° 校验让位给下方
                # 法兰级粗验收+MoveJ 微纠偏收口（终点仍回认证构型，护栏语义不降级）。
                # v14u：expect_target=段目标关节——目标锚定到位等待（上限 60s，每5s进度日志）。
                # v14w：净化只作用于发送关节；expect_target 仍是认证关节（到位判据不变）。
                # v14w37：位姿传递（动画=认证直线）+ flange_space 单位变换（校验/数字=法兰空间）。
                _send_pose = invH(robot.PoseFrame()) * robot.SolveFK(_send_q)
                _single_move_settle('MoveL', _send_pose, require_joints=False,
                                    expect_target=step['joints'], flange_space=True)
                try:
                    robot.setJoints(step['joints'])   # v14w39：模型钉到认证终点，清本地动画残留态
                except Exception:
                    pass
                # v14q：MovL 落点法兰级粗验收（≤8mm/≤1°）+ MoveJ 微纠偏收口（关节级 0.5° 罩终点）。
                # v14p 首航停在 0.95° 关节残差（法兰 4.61mm/0.616°）被 0.5° 护栏拦停——那是控制器
                # MovL 固有落点残差（v14l 5.5mm 双样本背书），不是构型错误；但终点必须回到认证构型，
                # 故验收通过后用一条短 MoveJ（~1° 关节差）收口，走 _single_move_settle 全套护栏。
                _actual, _is_static = _wait_controller_static(samples=3, interval=0.2)
                _mm, _deg = _movl_flange_accept(_actual, step['joints'])
                if _mm > MOVL_FLANGE_TOL_MM or _deg > MOVL_FLANGE_TOL_DEG:
                    raise RuntimeError('v14u 法兰级粗验收未过：停点法兰残差%.2fmm/%.2f°（容差%.1fmm/%.1f°），实测关节%s，停止待判读。'
                                       % (_mm, _deg, MOVL_FLANGE_TOL_MM, MOVL_FLANGE_TOL_DEG,
                                          ['%.2f' % v for v in _actual]))
                _jm = max(abs(a - b) for a, b in zip(_actual, step['joints']))
                if _jm > MOVE_OFFSET_TOL:
                    log(f"P{i}：v14u MovL 直发落点法兰级验收通过（残差{_mm:.2f}mm/{_deg:.2f}°），关节残差{_jm:.2f}°——发 MoveJ 微纠偏收口。")
                    _single_move_settle('MoveJ', step['joints'])
                _require_joints(step['joints'])
            elif (movl_direct and i in MOVL_DIRECT_BLOCK_POINTS and seg_mm is not None
                    and seg_mm <= MOVL_DIRECT_MAX_MM and seg_rot <= math.radians(0.5)):
                # ★ v14v4：本点被【禁直发名单】拦下 —— 明确告知，便于判读日志
                log(f"P{i}：⛔ 本点在【禁直发名单】MOVL_DIRECT_BLOCK_POINTS={MOVL_DIRECT_BLOCK_POINTS} 里 ⇒ "
                    f"不走法兰补偿直发，改走【细分途经点路径】（v14n 实测 17/17 通过、零事故的路径）。")
            elif waypoints:
                log(f"P{i}：执行预检方案 {step['method']}→MoveJ 细分，{len(waypoints)} 个途经点，终点关节={step['joints']}")
                for k, way in enumerate(waypoints, 1):
                    _move_with_completion_check('MoveJ', way, False)
                    _require_joints(way)
                _require_joints(step['joints'])
            else:
                log(f"P{i}：执行预检方案 {step['method']}，关节={step['joints']}")
                _move_with_completion_check(step['method'], step['joints'], split_moves)
                _require_joints(step['joints'])
            expected = step['joints']
            completed += 1
        log(f'实机执行完成：{completed}/{len(plan)}点。')
    except Exception as exc:
        log(f'实机任务停止，已完成{completed}点：{type(exc).__name__}: {exc}')
        if movl_direct and ('断连' in str(exc) or '未到位' in str(exc) or '落点偏差' in str(exc) or '粗验收' in str(exc)):
            log('【v14u】法兰补偿MOVL执行段出断连/落点指纹（v14w24 无勾选框；细分途经点路径保留在计划中，可作回退依据）。')
        try:
            actual, velocity, mode = _controller_feedback()
            log('停止时控制器实际反馈：关节=%s，速度=%s，模式=%s；不自动重发运动。' % (actual, velocity, mode))
        except Exception as feedback_error:
            log('停止时也无法取得控制器反馈：%s' % feedback_error)
    finally:
        _real_running = False
        try:
            _keepalive_stop.set()
            _ka_thread.join(timeout=3)
        except Exception:
            pass


def _point_to_segment_distance(p, a, b):
    """3D点到线段距离，单位mm。"""
    ax, ay, az = a
    bx, by, bz = b
    px, py, pz = p
    ab = (bx-ax, by-ay, bz-az)
    ap = (px-ax, py-ay, pz-az)
    ab2 = ab[0]*ab[0] + ab[1]*ab[1] + ab[2]*ab[2]
    if ab2 < 1e-12:
        return math.sqrt((px-ax)**2 + (py-ay)**2 + (pz-az)**2)
    t = (ap[0]*ab[0] + ap[1]*ab[1] + ap[2]*ab[2]) / ab2
    t = max(0.0, min(1.0, t))
    q = (ax+t*ab[0], ay+t*ab[1], az+t*ab[2])
    return math.sqrt((px-q[0])**2 + (py-q[1])**2 + (pz-q[2])**2)


def _tcp_position_from_joints(q):
    """关节角 -> 当前参考坐标系下的TCP位置，与轨迹输入使用同一坐标系。"""
    f = pose_to_fanuc_values(invH(robot.PoseFrame()) * robot.SolveFK(q) * robot.PoseTool())
    return (float(f[0]), float(f[1]), float(f[2]))


def _check_movej_tcp_trajectory(start_q, target_q, start_tcp_vals, target_tcp_vals, log, samples=30, max_deviation_mm=None):
    """
    在真正执行MoveJ之前，用关节空间线性插补采样，计算TCP轨迹相对
    起点-终点TCP直线段的最大偏离距离。

    目的：MoveL失败时，不再无条件MoveJ；只有MoveJ造成的TCP空间绕行
    没有超过允许值，才允许用MoveJ兜底。
    """
    if max_deviation_mm is None:
        max_deviation_mm = MOVEJ_FALLBACK_MAX_DEVIATION_MM

    start_q = [float(v) for v in start_q[:6]]
    target_q = [float(v) for v in target_q[:6]]
    a = (float(start_tcp_vals[0]), float(start_tcp_vals[1]), float(start_tcp_vals[2]))
    b = (float(target_tcp_vals[0]), float(target_tcp_vals[1]), float(target_tcp_vals[2]))

    log("开始检查 MoveJ 兜底轨迹：%d 个采样点，允许最大TCP偏离 %.3f mm" % (samples + 1, max_deviation_mm))
    max_dev = -1.0
    max_info = None

    for k in range(samples + 1):
        t = float(k) / float(samples)
        q = [start_q[j] + (target_q[j] - start_q[j]) * t for j in range(6)]
        try:
            p = _tcp_position_from_joints(q)
        except Exception as e:
            log("  MoveJ轨迹检查失败：第 %d/%d 个采样点 FK失败：%s: %s" % (k+1, samples+1, type(e).__name__, e))
            return False

        dev = _point_to_segment_distance(p, a, b)
        if dev > max_dev:
            max_dev = dev
            max_info = (k, t, q, p)

        if dev > max_deviation_mm:
            log("✕ MoveJ兜底轨迹拒绝：第 %d/%d 个采样点偏离TCP直线 %.3f mm > %.3f mm" %
                (k+1, samples+1, dev, max_deviation_mm))
            log("  t=%.3f  TCP=(%.3f, %.3f, %.3f)" % (t, p[0], p[1], p[2]))
            log("  因此不会执行这个MoveJ兜底动作，避免出现不可接受的大绕圈。")
            return False

    if max_info is not None:
        k, t, q, p = max_info
        log("✓ MoveJ兜底轨迹检查通过")
        log("  最大TCP偏离直线：%.3f mm（采样 %d/%d，t=%.3f）" % (max_dev, k+1, samples+1, t))
        log("  最大偏离点TCP=(%.3f, %.3f, %.3f)" % (p[0], p[1], p[2]))
    return True


# ============================================================
# 执行连续运动（MoveL失败时先检查MoveJ轨迹）
# ============================================================
def _collision_details():
    pairs = RDK.CollisionPairs()
    return '；'.join(f'{a.Name()}[连杆{ia}] 与 {b.Name()}[连杆{ib}]'
                    for a, b, ia, ib in pairs) or '路径碰撞或关节不可行'


def _enable_obstacle_checks():
    if RDK.RunMode() != RUNMODE_SIMULATE:
        raise RuntimeError('障碍物预检仅允许在仿真模式执行。')
    # 每次进入预检都清空预检缓存：缓存生命周期 = 单次预检规划，
    # 障碍物/工作站状态的变化在下一次预检即时生效。
    _plan_cache.clear()
    for name in ('安装台_650x650x80mm', '地面_禁止穿越', '磨砂圆柱_R150_H50', '挡板_半封闭3面'):
        obstacle = RDK.Item(name, ITEM_TYPE_OBJECT)
        if not obstacle.Valid():
            raise RuntimeError(f'缺少障碍物模型：{name}，请加载包含台子和地面的工作站。')
        if name == '安装台_650x650x80mm':
            if RDK.setCollisionActivePair(COLLISION_OFF, robot, obstacle, 0, 0) != 1:
                raise RuntimeError('无法配置安装台与固定底座的接触关系。')
        for link in range(1, 7):
            if RDK.setCollisionActivePair(COLLISION_ON, robot, obstacle, link, 0) != 1:
                raise RuntimeError(f'无法启用{name}与连杆{link}的碰撞检查。')
        tool_items = list(RDK.ItemList(ITEM_TYPE_TOOL))
        _handle = RDK.Item('门把手_bs1')   # v14w12：网格替换后可能为 OBJECT 类型，按名并入
        if _handle.Valid() and all(_handle.item != t.item for t in tool_items):
            tool_items.append(_handle)
        for tool in tool_items:
            parent = tool.Parent()
            while parent.Valid() and parent.item != robot.item:
                parent = parent.Parent()
            if parent.Valid() and RDK.setCollisionActivePair(COLLISION_ON, tool, obstacle) != 1:
                raise RuntimeError(f'无法启用{name}与工具的碰撞检查。')
    RDK.setCollisionActive(COLLISION_ON)


def _check_single_joint_path(end):
    _enable_obstacle_checks()
    saved = robot.Joints().list()[:6]
    try:
        RDK.Command('Trace', 'Off')
        RDK.Render(False)
        if _movej_test_cached(saved, end, 1) != 0:
            raise ValueError('单点MoveJ路径被拒绝：' + _collision_details())
    finally:
        robot.setJoints(saved)
        RDK.Render(True)


def _trajectory_pose(q):
    return invH(robot.PoseFrame()) * robot.SolveFK(q) * robot.PoseTool()


def _reorient_next_pose(records, i, rec):
    """v14w33：i 为 1-based 点号。若下一点存在且为【同 TCP 位姿纯换姿】（xyz 全同、姿态不同），
    返回下一点的 TCP 位姿 Mat，否则 None。用于换姿对的分支前视。"""
    try:
        if i >= len(records):
            return None
        nxt = records[i]          # 0-based 列表：下一条记录
        if nxt['type'] != 'TCP' or nxt.get('singular', False):
            return None
        va = [float(v) for v in rec['values'][:6]]
        vb = [float(v) for v in nxt['values'][:6]]
        if all(abs(va[k] - vb[k]) < 1e-9 for k in range(3)) and any(abs(va[k] - vb[k]) > 1e-9 for k in range(3, 6)):
            return fanuc_values_to_pose(*vb)
    except Exception:
        return None
    return None


def _linear_path_endpoint(start, target):
    """带结果缓存：分支重试时同一（起点, 目标）不重复计算。"""
    key = ('linear', _cache_key_joints(start), _cache_key_pose(target))
    if key in _plan_cache:
        return _plan_cache[key]
    result = _linear_path_endpoint_uncached(start, target)
    _plan_cache[key] = result
    return result


def _linear_path_endpoint_uncached(start, target):
    # 粗筛：10mm 采样点是 1mm 采样点的子集，粗筛失败则 1mm 细查必然失败，
    # 可直接拒绝；粗筛通过后再跑原有 1mm 细查，通过/拒绝判定与只跑 1mm 完全一致。
    status = robot.MoveL_Test(start, target, minstep_mm=10)
    if status == 0:
        status = robot.MoveL_Test(start, target, minstep_mm=1)
    if status != 0:
        return None, f'MoveL原生路径检查未通过（{status}）：' + _collision_details()
    # 本机MoveL_Test返回成功后Joints()可能为全零；从插补矩阵读取实际终点。
    # 碰撞判定已由上方同路径 1mm MoveL_Test 完成，此处仅提取终点关节，
    # 关闭碰撞检查提速（实测约快两个数量级）；整段权威碰撞复核仍在
    # _verify_obstacle_plan（碰撞开、1mm）进行。
    program = RDK.AddProgram('_TCP仿真_路径预检', robot)
    try:
        program.setVisible(False)
        robot.setJoints(start)
        program.setPoseFrame(robot.PoseFrame())
        program.setPoseTool(robot.PoseTool())
        program.MoveJ(start)
        program.MoveL(target)
        message, matrix, status = program.InstructionListJoints(mm_step=1, deg_step=1, collision_check=COLLISION_OFF)
        if status < 0:
            return None, message
        end = matrix.tr().rows[-1][:6]
        error_pose = invH(target) * _trajectory_pose(end)
        if norm(error_pose.Pos()) > .01 or pose_angle(error_pose) > math.radians(.01):
            raise RuntimeError('路径预检返回的终点不匹配目标TCP。')
        return end, message
    finally:
        program.Delete()


def _linear_waypoints(start, target, step_mm=None):
    """v13：从一条 MoveL 指令采样细分途经关节点（按 IK 顺序，无分支翻转）。

    用 InstructionListJoints(mm_step=LINEAR_SUBSTEP_MM, collision_check=COLLISION_OFF) 采样：
    途经点与 MoveL 执行的是同一条几何直线，且 IK 连续选解（避免用全局 SolveIK 时
    途经点在多解间跳变）。碰撞已由 _linear_path_endpoint 的 MoveL_Test@1mm 权威判定，
    此处不再重复。返回含终点的关节点列表；空列表表示采样失败（调用方回退直达）。"""
    if step_mm is None:
        step_mm = LINEAR_SUBSTEP_MM
    key = ('waypoints', _cache_key_joints(start), _cache_key_pose(target), round(float(step_mm), 3))
    if key in _plan_cache:
        return [q[:] for q in _plan_cache[key]]
    program = RDK.AddProgram('_TCP仿真_细分采样', robot)
    saved = robot.Joints().list()[:6]
    try:
        program.setVisible(False)
        robot.setJoints(start)
        program.setPoseFrame(robot.PoseFrame())
        program.setPoseTool(robot.PoseTool())
        program.MoveJ(start)
        program.MoveL(target)
        message, matrix, status = program.InstructionListJoints(mm_step=step_mm, deg_step=1, collision_check=COLLISION_OFF)
        cols = matrix.tr().rows if matrix is not None else []
        if status < 0 or not cols:
            return []
        # 丢弃比步长更密的重复点（InstructionListJoints 在奇异附近会加密采样）
        picked = [list(map(float, cols[0][:6]))]
        for row in cols[1:]:
            q = list(map(float, row[:6]))
            if max(abs(a - b) for a, b in zip(q, picked[-1])) >= step_mm / 10.0:
                picked.append(q)
        # 去尾：InstructionListJoints 可能带比目标多一点的收尾点，以关节距离最近的为准
        end_q, _ = _linear_path_endpoint(start, target)
        if end_q is not None and picked and max(abs(a - b) for a, b in zip(end_q, picked[-1])) > 1.0:
            picked[-1] = list(map(float, end_q))
        _plan_cache[key] = [q[:] for q in picked]
        return [q[:] for q in picked]
    finally:
        program.Delete()
        robot.setJoints(saved)


def _obstacle_posture_key(q, reference=None):
    table = RDK.Item('安装台_650x650x80mm', ITEM_TYPE_OBJECT)
    height = 0.0
    if table.Valid():
        elbow = invH(table.PoseAbs()) * robot.PoseAbs() * robot.JointPoses(q)[3]
        height = elbow.Pos()[2]
    return (-round(height, 6), sum((v-r)**2 for v, r in zip(q, reference or [0]*6)), tuple(q))


def _obstacle_joint_target(start, values, max_deviation=None, log=None):
    """带结果缓存：同一（起点, 目标, 偏离上限）的兜底选解不重复搜索。"""
    key = ('obstacle', _cache_key_joints(start), tuple(round(float(v), 6) for v in values[:6]),
           round(float(max_deviation), 6) if max_deviation is not None else None)
    if key in _plan_cache:
        cached = _plan_cache[key]
        if isinstance(cached, ValueError):
            raise cached
        return cached
    try:
        result = _obstacle_joint_target_uncached(start, values, max_deviation, log)
    except ValueError as exc:
        _plan_cache[key] = exc
        raise
    _plan_cache[key] = result
    return result


def _obstacle_joint_target_uncached(start, values, max_deviation=None, log=None):
    # v14-P2P：不再用 seed 候选/肘高排序，直接取离当前关节最近的逆解做逐级检查；
    # 最近解过不了偏离/碰撞时仍会在这里报错（单点 MoveJ 兜底路径保持可用）。
    lower, upper, _ = robot.JointLimits()
    candidates = [_nearest_ik_from_current(start, fanuc_to_pose(*values))]
    saved = robot.Joints().list()[:6]
    try:
        # 少量FK采样仅用于排序；不能替代后面的偏离复核与精细碰撞检查。
        a = _tcp_position_from_joints(start)
        table = RDK.Item('安装台_650x650x80mm', ITEM_TYPE_OBJECT)
        base_to_table = invH(table.PoseAbs()) * robot.PoseAbs()
        ranked = []
        for end in candidates:
            deviation, height = 0.0, float('inf')
            for k in range(11):
                q = [x + (y-x)*k/10 for x, y in zip(start, end)]
                deviation = max(deviation, _point_to_segment_distance(
                    _tcp_position_from_joints(q), a, values[:3]))
                height = min(height, (base_to_table * robot.JointPoses(q)[3]).Pos()[2])
            if max_deviation is not None and deviation > max_deviation:
                continue
            # 20mm一档，避免为很小的偏离差反复搜索；同档优先抬高肘部。
            ranked.append(((int(deviation/20), -height,
                            sum(abs(y-x) for x, y in zip(start, end))), end))
        checked = 0
        for _, end in sorted(ranked, key=lambda entry: entry[0]):
            if max_deviation is not None and not _check_movej_tcp_trajectory(
                    start, end, pose_to_fanuc_values(_trajectory_pose(start)), values,
                    lambda msg: None, samples=100, max_deviation_mm=max_deviation):
                continue
            checked += 1
            if _movej_test_cached(start, end, .25) == 0:
                if log is not None:
                    log(f'MoveJ快速筛选：{len(candidates)}个候选，{len(ranked)}个通过粗筛，精查{checked}条后找到合格路径。')
                return end
        raise ValueError('所有候选关节路径均碰撞、超出偏离限制或没有有效逆解。')
    finally:
        robot.setJoints(saved)


def _verify_obstacle_plan(start, plan):
    program = RDK.AddProgram('_TCP仿真_整段碰撞复核', robot)
    saved = robot.Joints().list()[:6]
    try:
        program.setVisible(False)
        program.setPoseFrame(robot.PoseFrame())
        program.setPoseTool(robot.PoseTool())
        program.MoveJ(start)
        for step in plan:
            for q in step['rewinds']:
                program.MoveJ(q)
            if step['method'] == 'MoveL' and not step.get('waypoints'):
                # v13 防呆：MoveL 步必须带细分途经点，否则规划层契约被破坏
                raise ValueError('整段碰撞复核：MoveL 步缺少细分途经点，拒绝。')
            getattr(program, step['method'])(step['joints'])
        message, matrix, status = program.InstructionListJoints(
            mm_step=1, deg_step=1, collision_check=COLLISION_ON)
        if status < 0 or 'collision' in message.lower():
            raise ValueError('整段碰撞复核未通过：' + message)
    finally:
        program.Delete()
        robot.setJoints(saved)


def _ik_branch_candidates(target_pose, reference):
    """v14c：某个 TCP 位姿的全部限位内 IK 分支（含 J6 圈数取近表示），
    与 _nearest_ik_from_current 同款筛选规则。"""
    solutions = robot.SolveIK_All(_tcp_target_to_flange(target_pose))
    lower, upper, _ = robot.JointLimits()
    lower, upper = lower.list(), upper.list()
    candidates = []
    for solution in solutions:
        q = [((float(v) + 180.0) % 360.0) - 180.0 for v in solution[:6]]
        if len(q) != 6:
            continue
        for turns6 in (0, -1, 1):
            candidate = q[:]
            candidate[5] += 360.0 * turns6
            if _real_limit_ok(candidate, lower, upper):
                if not any(max(abs(a-b) for a, b in zip(candidate, old)) < 1e-6 for old in candidates):
                    candidates.append(candidate)
    for q in candidates[:]:
        nearest = [min((v + 360*k for k in range(math.ceil((lower[j]-v)/360),
                       math.floor((upper[j]-v)/360)+1)), key=lambda a: abs(a-reference[j]))
                   for j, v in enumerate(q)]
        # v14w22：取近表示必须复核实机限位（此前漏检 ⇒ J1=193.59 混入实发被 -40001 拒）
        if not _real_limit_ok(nearest, lower, upper):
            continue
        if not any(max(abs(a-b) for a, b in zip(nearest, old)) < 1e-6 for old in candidates):
            candidates.append(nearest)
    return candidates


def _nearest_ik_from_current_lookahead(current_q, target_pose, lookahead_ok):
    """v14i：同 _nearest_ik_from_current，但要求选出的解能满足前视条件 lookahead_ok(cand)->bool；
    没有满足者时退回最近解（死路由后续救援链/种子重试兜底）。"""
    candidates = _ik_branch_candidates(target_pose, current_q)
    if not candidates:
        raise ValueError('没有限位内的逆解。')
    ranked = sorted(candidates, key=lambda q: sum((q[j]-current_q[j])**2 for j in range(6)))
    for cand in ranked:
        if lookahead_ok(cand):
            return cand[:]
    return ranked[0][:]


def _nearest_ik_from_current(current_q, target_pose):
    """v14-P2P：从全部逆解中选离当前关节角最近的解（含 J6 圈数取近）。

    与 test.py 的肘高排序不同：以【关节空间离当前构型最近】为准，相邻点之间不会突变构型。
    没有限位内解时抛 ValueError。"""
    solutions = robot.SolveIK_All(_tcp_target_to_flange(target_pose))
    lower, upper, _ = robot.JointLimits()
    lower, upper = lower.list(), upper.list()
    candidates = []
    for solution in solutions:
        q = [((float(v) + 180.0) % 360.0) - 180.0 for v in solution[:6]]
        if len(q) != 6:
            continue
        for turns6 in (0, -1, 1):
            candidate = q[:]
            candidate[5] += 360.0 * turns6
            if _real_limit_ok(candidate, lower, upper):
                if not any(max(abs(a-b) for a, b in zip(candidate, old)) < 1e-6 for old in candidates):
                    candidates.append(candidate)
    # 同一姿态再补一圈数取近的表示，避免强制归零导致大绕行。
    for q in candidates[:]:
        nearest = [min((v + 360*k for k in range(math.ceil((lower[j]-v)/360),
                       math.floor((upper[j]-v)/360)+1)), key=lambda a: abs(a-current_q[j]))
                   for j, v in enumerate(q)]
        # v14w22：取近表示必须复核实机限位（此前漏检 ⇒ J1=193.59 混入实发被 -40001 拒）
        if not _real_limit_ok(nearest, lower, upper):
            continue
        if not any(max(abs(a-b) for a, b in zip(nearest, old)) < 1e-6 for old in candidates):
            candidates.append(nearest)
    if not candidates:
        raise ValueError('没有限位内的逆解。')
    return min(candidates, key=lambda q: sum((q[j]-current_q[j])**2 for j in range(6)))[:]


def _checked_j6_rewinds(q, lower, upper, max_deviation):
    """返回可实际执行的整圈回绕列表（带缓存）；TCP空间偏离和碰撞都必须通过检查。"""
    key = ('rewinds', _cache_key_joints(q), tuple(round(float(v), 6) for v in lower[:6]),
           tuple(round(float(v), 6) for v in upper[:6]), round(float(max_deviation), 6))
    if key in _plan_cache:
        return [r[:] for r in _plan_cache[key]]
    results = []
    tcp = pose_to_fanuc_values(_trajectory_pose(q))
    for delta in (-360.0, 360.0):
        end = q[:]
        end[5] += delta
        if not lower[5] <= end[5] <= upper[5]:
            continue
        if not _check_movej_tcp_trajectory(q, end, tcp, tcp, lambda msg: None,
                                          samples=360, max_deviation_mm=max_deviation):
            continue
        if _movej_test_cached(q, end, 1) == 0:
            results.append(end)
    _plan_cache[key] = results
    return [r[:] for r in results]


def _plan_continuous_trajectory(records, max_deviation, log):
    """v14c：首点全分支种子枚举 + 整段重试。

    贪心最近解在换向步（如轨迹7 P6 的原地转 90°→180°）会把 wrist 构型选到贴圆柱，
    后续任何分支都碰；TCP仿真宏靠首点种子枚举+整段重试避开这类死路。v14c 移植该机制：
    种子按肘高排序优先，贪心只负责段内选解；某段死路（含 MoveL 兑底都失败）
    则整段换种子重试，全部种子失败才报错。"""
    _enable_obstacle_checks()
    if not math.isfinite(max_deviation) or max_deviation < 0:
        raise ValueError('MoveJ允许偏离必须是非负有限数。')
    for i, rec in enumerate(records):
        vals = rec['values']
        if rec['type'] not in ('TCP', 'JOINT') or len(vals) != 6 or not all(math.isfinite(v) for v in vals):
            raise ValueError(f'P{i+1}：点类型或六维数值无效。')
        if rec.get('singular', False):
            # v14a：恢复 v13 同款奇异点规则校验（P2P 规划层支持奇异点步）
            if rec['type'] != 'TCP' or i == 0 or records[i-1]['type'] != 'TCP' or records[i-1].get('singular', False):
                raise ValueError(f'P{i+1}：特异点必须紧跟普通TCP点。')
            if rec.get('spin360', False):
                if rec.get('j6_delta', 360) not in (-360, 360):
                    raise ValueError(f'P{i+1}：J6自转方向必须为+360或-360。')
                if max(abs(a - b) for a, b in zip(rec['values'], records[i-1]['values'])) > 1e-3:
                    raise ValueError(f'P{i+1}：J6自转360°特异点的六维数值必须与前一个TCP点完全相同。')
            elif rec.get('j6_delta', 180) not in (-180, 180):
                raise ValueError(f'P{i+1}：J6方向必须为+180或-180。')
    saved = robot.Joints().list()[:6]
    lower, upper, _ = robot.JointLimits()
    lower, upper = lower.list(), upper.list()
    # 先检查点本身可达，避免后面的不可达点触发整段分支重复搜索。
    unreachable = []
    for i, rec in enumerate(records, 1):
        if rec['type'] == 'TCP' and not rec.get('singular', False):
            target = fanuc_values_to_pose(*rec['values'])
            if robot.SolveIK_All(_tcp_target_to_flange(target)).size(1) == 0:
                unreachable.append(f'P{i}：没有逆解；' + _flange_target_description(target))
    if unreachable:
        raise ValueError('目标点不可达，尚未搜索连接路径：' + '；'.join(unreachable))
    if _movej_test_cached(saved, saved, 1) != 0:
        raise ValueError('起始姿态已碰撞，不能自动规划脱离：' + _collision_details())
    try:
        RDK.Render(False)
        # v14c：首点全分支种子枚举（肘高优先），某种子整段死路时换构型重试。
        first_tcp = next((r for r in records if r['type'] == 'TCP' and not r.get('singular', False)), None)
        if first_tcp is not None:
            seeds = _ik_branch_candidates(fanuc_values_to_pose(*first_tcp['values']), saved)
            seeds = [s for s in seeds if _movej_test_cached(saved, s, 1) == 0] or seeds
            seeds.sort(key=lambda s: _obstacle_posture_key(s, saved))
        else:
            seeds = [None]
        for seed_rank, seed in enumerate(seeds, 1):
            if len(seeds) > 1:
                log(f'—— 尝试首点分支种子 {seed_rank}/{len(seeds)}：' +
                    ('%s' % [round(v, 1) for v in seed] if seed else '无种子(关节轨迹)'))
            q = saved[:]
            plan = []
            try:
                seed_used = seed is None
                for i, rec in enumerate(records, 1):
                    rewinds = []
                    delta = None
                    method, fallback, waypoints = 'MoveJ', False, []
                    lookahead_ok = None  # v14j：循环顶初始化（首个TCP点走种子路径时前视绑定也可安全引用）
                    if rec['type'] == 'JOINT':
                        end = [float(v) for v in rec['values'][:6]]
                        note = '录入关节直达'
                    elif rec.get('singular', False):
                        # v14a：奇异点步——只转 J6（±180 换向 / ±360 自转）。
                        # ±180：从当前解纯转 J6，由下方 FK 校验把关；超限时先试反方向（终点位姿不变）再试整圈回绕。
                        target = fanuc_values_to_pose(*rec['values'])
                        delta = rec.get('j6_delta', 180)

                        def _fk_matches(candidate):
                            error_pose = invH(target) * _trajectory_pose(candidate)
                            return norm(error_pose.Pos()) <= 1e-3 and pose_angle(error_pose) <= math.radians(.01)

                        end = q[:]
                        end[5] += delta
                        if not lower[5] <= end[5] <= upper[5]:
                            alt = q[:]
                            alt[5] -= delta
                            if lower[5] <= alt[5] <= upper[5]:
                                log(f'P{i}：J6 {delta:+d}°超限，改用反方向 {-delta:+d}°（终点位姿不变）。')
                                end, delta = alt, -delta
                            if not lower[5] <= end[5] <= upper[5]:
                                for rewound in _checked_j6_rewinds(q, lower, upper, max_deviation):
                                    if lower[5] <= rewound[5] + delta <= upper[5]:
                                        rewinds.append(rewound[:])
                                        q = rewound
                                        end = q[:]
                                        end[5] += delta
                                        break
                                else:
                                    raise ValueError(f'P{i}：J6 {delta:+d}°超限：反方向与整圈回绕均不可行。')
                        if not _fk_matches(end):
                            raise ValueError(f'P{i}：仅旋转J6无法到达所标注TCP，请检查特异点标记/工具。')
                        # v14d：换向步碰撞时，先试反方向（终点位姿不变），再试整圈回绕——
                        # TCP仿真靠方向枚举能避开这类碰撞，P2P 此前只在超限时才换向。
                        # v14j：反方向终点=当前解−delta（旧代码误算 q−2δ，朝向未翻转、FK 必不匹配，
                        # 15/15 种子全死于此——probe_p14_lookahead.py 坐实）。
                        if _movej_test_cached(q, end, 1) != 0:
                            alt = q[:]
                            alt[5] -= delta
                            flipped = False
                            if lower[5] <= alt[5] <= upper[5] and _fk_matches(alt) and _movej_test_cached(q, alt, 1) == 0:
                                log(f'P{i}：J6 {delta:+d}°扫过障碍，改用反方向 {-delta:+d}°（终点位姿不变）。')
                                end, delta, flipped = alt, -delta, True
                            if not flipped:
                                for rewound in _checked_j6_rewinds(q, lower, upper, max_deviation):
                                    cand = rewound[:]
                                    cand[5] += delta
                                    if lower[5] <= cand[5] <= upper[5] and _fk_matches(cand) and _movej_test_cached(q, cand, 1) == 0:
                                        log(f'P{i}：J6 {delta:+d}°两方向均碰，先整圈回绕再换向。')
                                        rewinds.append(rewound[:])
                                        q, end, flipped = rewound, cand, True
                                        break
                            if not flipped:
                                # v14f：两方向都碰——先切到同位姿的其他 IK 分支（碰撞预检过），
                                # 从那里再换向；途经的构型跳记入 rewinds 由执行层逐跳执行。
                                # v14j：枚举基准改为当前（未翻转）位姿——旧代码误用翻转后 target，
                                # 候选再 ±180 回到未翻转位姿，FK 对 target 永不匹配，结构性必死。
                                for cand in sorted(_ik_branch_candidates(_trajectory_pose(q), q),
                                                   key=lambda c: sum((c[j]-q[j])**2 for j in range(6))):
                                    for sgn in (delta, -delta):
                                        after = cand[:]
                                        after[5] += sgn
                                        if not (lower[5] <= after[5] <= upper[5] and _fk_matches(after)):
                                            continue
                                        if _movej_test_cached(q, cand, 1) == 0 and _movej_test_cached(cand, after, 1) == 0:
                                            log(f'P{i}：J6 ±180°两方向均碰，先切IK分支再换向（rewinds 跳转）。')
                                            rewinds.append(cand[:])
                                            q, end, delta, flipped = cand, after, sgn, True
                                            break
                                    if flipped:
                                        break
                            if not flipped:
                                # v14g：同位姿先 MoveL 到场再换向——MoveL 连续选解给出的构型
                                # 正是 TCP仿真 实测可换向的构型（贪心最近解构型两方向都扫障碍）。
                                lin_end, lin_detail = _linear_path_endpoint(q, target)
                                if lin_end is not None:
                                    pre_waypoints = _linear_waypoints(q, target)
                                    if pre_waypoints:
                                        for sgn in (delta, -delta):
                                            after = lin_end[:]
                                            after[5] += sgn
                                            if not (lower[5] <= after[5] <= upper[5] and _fk_matches(after)):
                                                continue
                                            if _movej_test_cached(lin_end, after, 1) == 0:
                                                log(f'P{i}：J6 两方向均碰，先 MoveL 到场（连续选解构型）再{sgn:+d}°换向。')
                                                plan.append(dict(method='MoveL', joints=lin_end[:], special=False,
                                                                 fallback=False, rewinds=[], j6_delta=None,
                                                                 waypoints=pre_waypoints, p2p_note='换向前MoveL到场'))
                                                q, end, delta, flipped = lin_end[:], after, sgn, True
                                                break
                            if not flipped:
                                raise ValueError(f'P{i}：J6 ±180°换向两方向均碰撞（含回绕/分支/MoveL到场尝试），该构型不可行。')
                        note = ('J6自转%+d°' % delta) if rec.get('spin360', False) else ('J6换向%+d°' % delta)
                    else:
                        target = fanuc_values_to_pose(*rec['values'])
                        # v14h：与前一点同位姿（停顿点，如轨迹7 P7）——不重新选解，
                        # 保持当前构型不动，只往计划里记一个停顿点。
                        if max(abs(_trajectory_pose(q).Pos()[j] - target.Pos()[j]) for j in range(3)) < 1e-3 and \
                           pose_angle(invH(target) * _trajectory_pose(q)) < math.radians(.01):
                            plan.append(dict(method='MoveJ', joints=q[:], special=False, fallback=False,
                                             rewinds=[], j6_delta=None, waypoints=[], p2p_note='同位姿停顿'))
                            continue
                        if not seed_used:
                            end = seed[:]  # v14c：首个TCP点直接采用种子分支（离起点可达性已在种子筛选时验证）
                            seed_used = True
                        else:
                            # v14i：前视——下一个执行点是 ±180 换向时，本点选解必须能完成那次换向
                            #（两方向任一可通行），否则贪心构型会把换向逼成死路。
                            nxt = records[i] if i < len(records) else None
                            lookahead_ok = None
                            if nxt is not None and nxt.get('singular', False) and not nxt.get('spin360', False):
                                nxt_values = nxt['values']
                                def lookahead_ok(cand, _vals=nxt_values, _lower=lower, _upper=upper):
                                    nxt_target = fanuc_values_to_pose(*_vals)
                                    for sgn in (180, -180):
                                        after = cand[:]
                                        after[5] += sgn
                                        if not (_lower[5] <= after[5] <= _upper[5]):
                                            continue
                                        err = invH(nxt_target) * _trajectory_pose(after)
                                        if norm(err.Pos()) > 1e-3 or pose_angle(err) > math.radians(.01):
                                            continue
                                        if _movej_test_cached(cand, after, 1) == 0:
                                            return True
                                    return False
                                log(f'P{i}：前视模式（P{i+1}为±180换向，选解需兼顾换向可行性）。')
                            end = (_nearest_ik_from_current_lookahead(q, target, lookahead_ok)
                                   if lookahead_ok else _nearest_ik_from_current(q, target))
                        note = 'TCP最近解直达'
                        forced_lin = False
                        # v14w24：短直线工作段强制 MoveL——P2→P3 这类 ≤210mm/姿态恒定 的
                        # 贴面平移，工艺不允许 MoveJ 关节弧绕行，直走直线（判据与直发门禁同款）。
                        # 前视夜（下一点±180换向）：直线末端同样具备换向资格才强制，否则回落
                        # MoveJ 前视绑定（保住换向可行性纪律）。
                        _rel = _trajectory_pose(q) * invH(target)
                        _seg_mm_f = norm(_rel.Pos())
                        _force_ok = _seg_mm_f <= MOVL_DIRECT_MAX_MM and pose_angle(_rel) <= math.radians(0.5)
                        # v14w33c：回撤段（TCP y 朝基座 >10mm）且下一点是同位姿换姿 ⇒ 让位 MoveJ
                        # 分支前视（强制 MoveL 的端点分支由直线 IK 连续性锁死，会对下一点无路：
                        # P5→P6→P7 实录 P7 被迫 49 跳细分）。工艺贴面滑移（Δy≈0）不受影响。
                        if _force_ok and i >= 2 and _reorient_next_pose(records, i, rec) is not None:
                            try:
                                _y_prev = float(records[i - 2]['values'][1])
                                if float(rec['values'][1]) - _y_prev > 10.0:
                                    _force_ok = False
                                    log(f'P{i}：回撤段且下一点为同位姿换姿——短直线让位 MoveJ 分支前视（v14w33c）。')
                            except Exception:
                                pass
                        if _force_ok:
                            lin_end_f, lin_detail_f = _linear_path_endpoint(q, target)
                            _lin_ok_f = (lin_end_f is not None
                                         and not _real_interfere_combo(lin_end_f)   # v14w26 组合禁区
                                         and (lookahead_ok is None or lookahead_ok(lin_end_f)))
                            if _lin_ok_f:
                                waypoints = _linear_waypoints(q, target)
                                if waypoints:
                                    end, method, fallback = lin_end_f, 'MoveL', True
                                    note = '短直线强制MoveL'
                                    forced_lin = True
                                    log(f'P{i}：短直线段（{_seg_mm_f:.1f}mm/姿态恒定）按工艺直走 MoveL（不尝试 MoveJ 弧）。')
                            elif lin_end_f is not None:
                                log(f'P{i}：短直线段直线末端无前视换向资格，回落 MoveJ 前视绑定。')
                            else:
                                log(f'P{i}：短直线段 MoveL 不可通行（{lin_detail_f}），回落 MoveJ 尝试。')
                        bound_applied = False
                        # v14j：前视绑定执行——本点是换向前夜：前视选出的构型若弧碰，不得退 MoveL
                        # （连续选解会静默锁回当前族，把死局推迟到换向步才爆——种子13 实证），
                        # 也不得由 v14c 救援收无前视资格的分支；只能换用其他前视合格分支直达，
                        # 全部失败则本构型判死、整段换种子重试。
                        if not forced_lin and lookahead_ok is not None and _movej_test_cached(q, end, 1) != 0:
                            detail_bound = _collision_details()
                            bound = None
                            for cand in sorted(_ik_branch_candidates(target, q),
                                               key=lambda c: sum((c[j]-q[j])**2 for j in range(6))):
                                if lookahead_ok(cand) and _movej_test_cached(q, cand, 1) == 0:
                                    bound = cand
                                    break
                            if bound is not None:
                                end, note, bound_applied = bound[:], '前视绑定避障直达', True
                                log(f'P{i}：前视构型弧碰（{detail_bound}），改用另一前视合格分支直达（前视绑定）。')
                            else:
                                raise ValueError(f'P{i}：MoveJ弧碰撞（{detail_bound}），其余前视合格分支均不可通行；'
                                                 '拒绝退 MoveL（连续选解会丢前视资格），本构型判死。')
                        # v14b：MoveJ 直达弧碰撞时，退回 v13 验证过的 MoveL 直线细分执行。
                        # v14w24：强制 MoveL 段不再尝试/回退 MoveJ（工艺直线优先）。
                        if not forced_lin and not bound_applied and _movej_test_cached(q, end, 1) != 0:
                            detail = _collision_details()
                            lin_end, lin_detail = _linear_path_endpoint(q, target)
                            if lin_end is None:
                                # v14c：直线也碰——枚举该目标全部 IK 分支找可通行 MoveJ（换构型救援）
                                # v14w33b：若下一点是【同位姿纯换姿】，优先选「下一点也能单条 MoveJ 贯通」
                                # 的救援分支（P6→P7 教训：P6 为自避碰选的分支对 P7 无路 ⇒ 49 跳细分拖死执行）。
                                _cands = sorted(_ik_branch_candidates(target, q),
                                                key=lambda c: sum((c[j] - q[j]) ** 2 for j in range(6)))
                                _nxt_pose = None
                                try:
                                    if i < len(records):
                                        _nr = records[i]
                                        if _nr['type'] == 'TCP' and not _nr.get('singular', False):
                                            _va = [float(v) for v in rec['values'][:6]]
                                            _vb = [float(v) for v in _nr['values'][:6]]
                                            if (all(abs(_va[k] - _vb[k]) < 1e-9 for k in range(3))
                                                    and any(abs(_va[k] - _vb[k]) > 1e-9 for k in range(3, 6))):
                                                _nxt_pose = fanuc_values_to_pose(*_nr['values'][:6])
                                except Exception:
                                    _nxt_pose = None
                                rescued = None
                                if _nxt_pose is not None:
                                    for cand in _cands:
                                        if _movej_test_cached(q, cand, 1) != 0:
                                            continue
                                        _ok_nxt = False
                                        for nb in _ik_branch_candidates(_nxt_pose, cand):
                                            if (_real_limit_ok(nb, lower, upper)
                                                    and not _real_interfere_combo(nb)
                                                    and _movej_test_cached(cand, nb, 1) == 0):
                                                _ok_nxt = True
                                                break
                                        if _ok_nxt:
                                            rescued = cand
                                            log(f'P{i}：下一点为同位姿换姿——救援分支带前视，选可与下一点单条 MoveJ 贯通的分支。')
                                            break
                                if rescued is None:
                                    for cand in _cands:
                                        if _movej_test_cached(q, cand, 1) == 0:
                                            rescued = cand
                                            break
                                if rescued is None:
                                    raise ValueError(f'P{i}：MoveJ弧碰撞（{detail}），且MoveL直线也失败：{lin_detail}；'
                                                     '该目标全部IK分支均不可通行。')
                                end, note = rescued[:], 'IK分支救援直达'
                                log(f'P{i}：最近解与直线均碰，切换IK分支救援成功。')
                            else:
                                # v14w33：同位姿/近零长（≤1mm）纯换姿段——MoveL 细分会把 90° 姿态差
                                # 切成数十跳小 MoveJ（10-21 P6→P7 实录 49 跳×每跳断连周期≈3s，
                                # 拖死执行）。优先搜无碰 MoveJ 分支单条直达（分支连续性绑死时
                                # 最近解弧碰≠无解）；搜不到再落回 MoveL 细分兜底。
                                # v14w34：_seg_mm_ro 必须是真实位置差——相对位姿平移模长在原地换姿
                                # 时被旋转杠杆放大（p−R·p，(0,-650,380) 处 90° 即 1064.8mm），
                                # 旧算式使 ≤1mm 门槛从未成立、两个搜索入口从未触发。
                                _pa = _trajectory_pose(q).Pos()
                                _pb = target.Pos()
                                _seg_mm_ro = math.sqrt(sum((_pa[_k] - _pb[_k]) ** 2 for _k in range(3)))
                                reorient_direct = None
                                if _seg_mm_ro <= 1.0:
                                    for cand in sorted(_ik_branch_candidates(target, q),
                                                       key=lambda c: sum((c[j]-q[j])**2 for j in range(6))):
                                        if (not _real_interfere_combo(cand)
                                                and _real_limit_ok(cand, lower, upper)
                                                and (lookahead_ok is None or lookahead_ok(cand))
                                                and _movej_test_cached(q, cand, 1) == 0):
                                            reorient_direct = cand
                                            break
                                if reorient_direct is not None:
                                    end, note = reorient_direct[:], '同位姿换姿MoveJ直达'
                                    method, fallback = 'MoveJ', False
                                    waypoints = []
                                    log(f'P{i}：同位姿换姿——MoveL 细分会碎成数十小段，改用无碰 MoveJ 分支单条直达。')
                                elif _seg_mm_ro <= 1.0 and plan and rec['type'] == 'TCP' and i >= 2:
                                    # v14w33d：回改上一步（已入计划、未执行）为可与本点单条 MoveJ 贯通的
                                    # 分支——上一步若走最近解直达/救援，其分支未必对本点有路（P6→P7 实录）。
                                    # 改关节目标后两跳路径均当场重检，证书完整。
                                    _prev_step = plan[-1]
                                    _prev_q = _prev_step['joints']
                                    _prev_prev = plan[-2]['joints'] if len(plan) >= 2 else saved
                                    _prev_pose = fanuc_values_to_pose(*records[i - 2]['values'][:6])
                                    reorient_direct = None
                                    for c6 in sorted(_ik_branch_candidates(_prev_pose, _prev_prev),
                                                     key=lambda c: sum((c[k] - _prev_q[k]) ** 2 for k in range(6))):
                                        if _real_interfere_combo(c6) or not _real_limit_ok(c6, lower, upper):
                                            continue
                                        if _movej_test_cached(_prev_prev, c6, 1) != 0:
                                            continue
                                        for c7 in sorted(_ik_branch_candidates(target, c6),
                                                         key=lambda c: sum((c[k] - c6[k]) ** 2 for k in range(6))):
                                            if _real_interfere_combo(c7) or not _real_limit_ok(c7, lower, upper):
                                                continue
                                            if lookahead_ok is not None and not lookahead_ok(c7):
                                                continue
                                            if _movej_test_cached(c6, c7, 1) != 0:
                                                continue
                                            _prev_step['joints'] = c6[:]
                                            reorient_direct = c7
                                            break
                                        if reorient_direct is not None:
                                            break
                                    if reorient_direct is not None:
                                        end, note = reorient_direct[:], '同位姿换姿MoveJ直达'
                                        method, fallback = 'MoveJ', False
                                        waypoints = []
                                        log(f'P{i}：回改上一步分支后，本点取得单条 MoveJ 直达（两跳均重检无碰）。')
                                if reorient_direct is not None:
                                    pass   # 已在上方处理
                                else:
                                    waypoints = _linear_waypoints(q, target)
                                    if not waypoints:
                                        raise ValueError(f'P{i}：MoveJ弧碰撞（{detail}），MoveL细分采样失败，拒绝。')
                                    end, method, fallback = lin_end, 'MoveL', True
                                    note = 'MoveJ弧碰退回MoveL细分'
                                    log(f'P{i}：MoveJ弧碰撞（{detail}），改走 MoveL 直线细分（{len(waypoints)} 途经点）。')
                    if not all(lower[j] <= end[j] <= upper[j] for j in range(6)):
                        raise ValueError(f'P{i}：关节超限，J6目标={end[5]:.3f}°。')
                    if method == 'MoveJ' and _movej_test_cached(q, end, 1) != 0:
                        # v14e：普通TCP点最后一级救援——v13 遗产 _obstacle_joint_target
                        # （21候选、肘高排序、限TCP偏离）选避障构型，TCP仿真靠它在同一站过关。
                        try:
                            end = _obstacle_joint_target(q, rec['values'], max_deviation, log)
                            note = '避障选解直达'
                        except ValueError:
                            raise ValueError(f'P{i}：MoveJ路径检查失败（含避障选解）：' + _collision_details())
                        if _movej_test_cached(q, end, 1) != 0:
                            raise ValueError(f'P{i}：MoveJ路径检查失败：' + _collision_details())
                    # v14w25：J6 恰=±360 边界值被控制器 -40006 拒收（10-15 17:26/17:33 实录）。
                    # v14w32：±359.999 内推仍防不住「J6 单轴被丢弃」（10-21 P4 实证：J1~J5 全到、
                    # J6 纹丝停在 180、误差 180°）——改为换 (−180,180] 同角表示（359.999→−0.001），
                    # J6 彻底离开 ±360 邻域。换表示会翻转 MoveJ 弧方向 ⇒ 必须重检路径，不过即报规划错误。
                    # spin360/多圈值（|J6|>360.001）不在此列，防绞坏自转语义。
                    if abs(end[5]) >= 359.999 and abs(end[5]) <= 360.001 and not rec.get('spin360'):
                        _j6n = end[5] - math.copysign(360.0, end[5])
                        log(f'P{i}：J6={end[5]:.3f}° 贴 ±360 边界，换同角表示 {_j6n:.3f}°（v14w32：±359.999 仍被丢轴，彻底离开边界邻域）。')
                        end[5] = _j6n
                        for _wp in waypoints:
                            if abs(_wp[5]) >= 359.999 and abs(_wp[5]) <= 360.001:
                                _wp[5] = _wp[5] - math.copysign(360.0, _wp[5])
                        if method == 'MoveJ' and _movej_test_cached(q, end, 1) != 0:
                            raise ValueError(f'P{i}：J6 换同角表示后 MoveJ 路径碰撞：' + _collision_details())
                    # v14w26：解落入实机自干涉组合区（J4×J5，-40006）——MoveJ 解自动换无碰安全
                    # 分支直达；直线段落区（强制/兜底）整段换种子；无安全分支则判死。
                    if _real_interfere_combo(end):
                        if method == 'MoveJ' and rec['type'] == 'TCP' and not rec.get('singular', False):
                            rescued_if = None
                            for cand_if in sorted(_ik_branch_candidates(target, q),
                                                   key=lambda c: sum((c[j]-q[j])**2 for j in range(6))):
                                if (_real_limit_ok(cand_if, lower, upper)
                                        and not _real_interfere_combo(cand_if)
                                        and _movej_test_cached(q, cand_if, 1) == 0):
                                    rescued_if = cand_if
                                    break
                            if rescued_if is None:
                                raise ValueError(f'P{i}：全部无碰分支均落入实机自干涉组合区'
                                                 f'（|J4|>{REAL_INTERFERE_J4_MAX:.0f} 且 |J5|>{REAL_INTERFERE_J5_MIN:.0f}，-40006 实录区），本构型判死。')
                            log(f'P{i}：预选解落入实机自干涉组合区（J4={end[3]:.1f}°, J5={end[4]:.1f}°），换安全分支直达。')
                            end = rescued_if[:]
                            note = '自干涉安全分支直达'
                        else:
                            raise ValueError(f'P{i}：该步解落入实机自干涉组合区（J4={end[3]:.1f}°, J5={end[4]:.1f}°），换种子重试。')
                    plan.append(dict(method=method, joints=end[:], special=rec.get('singular', False), fallback=False,
                                     rewinds=rewinds, j6_delta=delta,
                                     waypoints=waypoints, p2p_note=note))
                    q = end[:]
                _verify_obstacle_plan(saved, plan)
                log(f'P2P+奇异点整段路径预检通过：{len(plan)}点。')
                return plan
            except ValueError as exc:
                if seed_rank >= len(seeds):
                    raise
                log(f'种子 {seed_rank}/{len(seeds)} 在此构型失败（{exc}），换下一构型整段重试…')
    finally:
        robot.setJoints(saved)
        RDK.Render(True)

root = tk.Tk()
root.title("RoboDK - 机械臂运动控制（P2P v14w41）")
root.geometry("1200x750")
root.resizable(True, True)

tk.Label(root, text="Dobot CR5 运动控制", font=("Microsoft YaHei", 16, "bold")).pack(pady=10)

notebook = ttk.Notebook(root)
notebook.pack(fill=tk.BOTH, expand=True, padx=10, pady=5)

# ---- 选项卡 1：单点运动 ----
tab_single = ttk.Frame(notebook)
notebook.add(tab_single, text="单点运动")

frame_coord = tk.LabelFrame(tab_single, text="目标 TCP（Fanuc 格式）")
frame_coord.pack(fill=tk.X, padx=10, pady=10)

names = ["X (mm)", "Y (mm)", "Z (mm)", "Rx (deg)", "Ry (deg)", "Rz (deg)"]
defaults = ["0.000", "-241.500", "1047.000", "-90.000", "0.000", "180.000"]
entries_single = []

for i in range(6):
    tk.Label(frame_coord, text=names[i]).grid(row=0, column=i*2, padx=5, pady=10)
    e = tk.Entry(frame_coord, width=12)
    e.insert(0, defaults[i])
    e.grid(row=0, column=i*2+1, padx=5, pady=10)
    entries_single.append(e)

frame_mtype = tk.Frame(tab_single)
frame_mtype.pack(fill=tk.X, padx=10, pady=5)
move_type = tk.StringVar(value="MoveL")
tk.Radiobutton(frame_mtype, text="MoveL (直线)", variable=move_type, value="MoveL").pack(side=tk.LEFT, padx=10)
tk.Radiobutton(frame_mtype, text="MoveJ (关节)", variable=move_type, value="MoveJ").pack(side=tk.LEFT, padx=10)

btn_single_frame = tk.Frame(tab_single)
btn_single_frame.pack(fill=tk.X, padx=10, pady=5)

def _read_current():
    read_current(entries_single)
def _fill_current():
    fill_current(entries_single)
def _check_ik():
    check_ik_single(entries_single)
def _exec_single():
    execute_single(entries_single, move_type.get())

tk.Button(btn_single_frame, text="读取当前 TCP", command=_read_current, width=15).pack(side=tk.LEFT, padx=3)
tk.Button(btn_single_frame, text="当前 TCP -> 输入框", command=_fill_current, width=20).pack(side=tk.LEFT, padx=3)
tk.Button(btn_single_frame, text="检测可达性", command=_check_ik, width=15, bg="#2196F3", fg="white").pack(side=tk.LEFT, padx=3)
tk.Button(btn_single_frame, text="执行运动", command=_exec_single, width=20,
          font=("Microsoft YaHei", 10, "bold"), bg="#4CAF50", fg="white").pack(side=tk.LEFT, padx=3)


# ---- 选项卡 2：目标关节运动（实机） ----
tab_joint = ttk.Frame(notebook)
notebook.add(tab_joint, text="目标关节运动")

frame_joint = tk.LabelFrame(tab_joint, text="目标关节（deg）")
frame_joint.pack(fill=tk.X, padx=10, pady=10)

joint_names = ["J1 (deg)", "J2 (deg)", "J3 (deg)", "J4 (deg)", "J5 (deg)", "J6 (deg)"]
joint_defaults = ["0.000", "0.000", "0.000", "0.000", "0.000", "0.000"]
entries_joint = []

for i in range(6):
    tk.Label(frame_joint, text=joint_names[i]).grid(row=0, column=i*2, padx=5, pady=10)
    e = tk.Entry(frame_joint, width=12)
    e.insert(0, joint_defaults[i])
    e.grid(row=0, column=i*2+1, padx=5, pady=10)
    entries_joint.append(e)

btn_joint_frame = tk.Frame(tab_joint)
btn_joint_frame.pack(fill=tk.X, padx=10, pady=8)

def _read_current_joint_values():
    read_current_joints(entries_joint)

def _fill_current_joints():
    fill_current_joints(entries_joint)

def _exec_joint():
    execute_joint_target(entries_joint)

def _zero_joints():
    clear_joint_target(entries_joint)

tk.Button(btn_joint_frame, text="读取当前关节", command=_read_current_joint_values, width=14).pack(side=tk.LEFT, padx=3)
tk.Button(btn_joint_frame, text="当前关节 -> 输入框", command=_fill_current_joints, width=20).pack(side=tk.LEFT, padx=3)
tk.Button(btn_joint_frame, text="执行指定关节 MoveJ", command=_exec_joint, width=24,
          font=("Microsoft YaHei", 10, "bold"), bg="#FF9800", fg="white").pack(side=tk.LEFT, padx=3)
tk.Button(btn_joint_frame, text="清零", command=_zero_joints, width=10).pack(side=tk.LEFT, padx=3)

tk.Label(tab_joint,
         text="输入 J1~J6 目标角度（deg）；完整关节路径预检通过后才发送实机 MoveJ。",
         fg="#555555").pack(anchor=tk.W, padx=15, pady=5)
tk.Label(tab_joint,
         text="安全提示：首次测试建议只改变一个关节、改变 5~10°，确认方向和角度定义正确后再进行大角度运动。",
         fg="#C62828").pack(anchor=tk.W, padx=15, pady=2)

# ---- 选项卡 3：连续运动 ----
tab_traj = ttk.Frame(notebook)
notebook.add(tab_traj, text="连续运动")

frame_traj_input = tk.LabelFrame(
    tab_traj,
    text="连续运动点输入：每次输入 1 个 TCP 点或 1 组关节角度，点击“检查并加入”"
)
frame_traj_input.pack(fill=tk.X, padx=10, pady=10)

type_frame = tk.Frame(frame_traj_input)
type_frame.pack(fill=tk.X, padx=8, pady=5)

tk.Label(type_frame, text="点类型：").pack(side=tk.LEFT, padx=3)

traj_type = tk.StringVar(value="TCP")
tk.Radiobutton(
    type_frame, text="TCP（X,Y,Z,Rx,Ry,Rz）",
    variable=traj_type, value="TCP"
).pack(side=tk.LEFT, padx=8)

tk.Radiobutton(
    type_frame, text="关节（J1~J6）",
    variable=traj_type, value="JOINT"
).pack(side=tk.LEFT, padx=8)

traj_names_tcp = ["X", "Y", "Z", "Rx", "Ry", "Rz"]
traj_names_joint = ["J1", "J2", "J3", "J4", "J5", "J6"]

traj_entries = []

# ---- 末端特异点设置 ----
singular_var = tk.BooleanVar(value=False)
j6_direction_var = tk.IntVar(value=180)

singular_frame = tk.Frame(frame_traj_input)
singular_frame.pack(fill=tk.X, padx=8, pady=3)

tk.Checkbutton(
    singular_frame,
    text="末端特异点（跳过IK，仅J6转动）",
    variable=singular_var
).pack(side=tk.LEFT, padx=3)

tk.Label(singular_frame, text="J6方向：").pack(side=tk.LEFT, padx=(15, 3))
tk.Radiobutton(singular_frame, text="+180°", variable=j6_direction_var, value=180).pack(side=tk.LEFT, padx=3)
tk.Radiobutton(singular_frame, text="-180°", variable=j6_direction_var, value=-180).pack(side=tk.LEFT, padx=3)
spin_var = tk.BooleanVar(value=False)
tk.Checkbutton(singular_frame, text="J6自转360°（第二类，六维与前点相同）", variable=spin_var).pack(side=tk.LEFT, padx=3)

# 输入框单独放在 grid 子容器中。
# frame_traj_input 本身使用 pack 管理子控件，不能再直接对它的子控件使用 grid。
traj_value_frame = tk.Frame(frame_traj_input)
traj_value_frame.pack(fill=tk.X, padx=8, pady=5)

for i in range(6):
    tk.Label(
        traj_value_frame,
        text=traj_names_tcp[i]
    ).grid(row=0, column=i * 2, padx=3, pady=8)

    e = tk.Entry(traj_value_frame, width=12)
    e.grid(row=0, column=i * 2 + 1, padx=4, pady=8)
    traj_entries.append(e)

# 默认先按 TCP 输入显示
tcp_defaults = ["0.000", "-241.500", "1047.000", "-90.000", "0.000", "180.000"]
for e, val in zip(traj_entries, tcp_defaults):
    e.insert(0, val)


def _update_traj_labels_and_defaults():
    """切换 TCP/关节输入时，更新标签和默认值。"""
    names = traj_names_tcp if traj_type.get() == "TCP" else traj_names_joint
    defaults = (
        tcp_defaults
        if traj_type.get() == "TCP"
        else ["0.000"] * 6
    )

    for i, e in enumerate(traj_entries):
        # grid 上的 Label 位于当前列
        for widget in traj_value_frame.grid_slaves(row=0, column=i * 2):
            widget.configure(text=names[i])

        e.delete(0, tk.END)
        e.insert(0, defaults[i])


tk.Radiobutton(
    type_frame, text="TCP（X,Y,Z,Rx,Ry,Rz）",
    variable=traj_type, value="TCP",
    command=_update_traj_labels_and_defaults
).pack_forget()

# 重新建立带 command 的两个单选按钮
for widget in list(type_frame.pack_slaves()):
    if isinstance(widget, tk.Radiobutton):
        widget.destroy()

tk.Radiobutton(
    type_frame, text="TCP（X,Y,Z,Rx,Ry,Rz）",
    variable=traj_type, value="TCP",
    command=_update_traj_labels_and_defaults
).pack(side=tk.LEFT, padx=8)

tk.Radiobutton(
    type_frame, text="关节（J1~J6）",
    variable=traj_type, value="JOINT",
    command=_update_traj_labels_and_defaults
).pack(side=tk.LEFT, padx=8)

btn_traj_input = tk.Frame(tab_traj)
btn_traj_input.pack(fill=tk.X, padx=10, pady=3)

tk.Button(
    btn_traj_input,
    text="检查并加入当前点",
    command=add_and_check_trajectory_point,
    width=22,
    bg="#2196F3",
    fg="white",
    font=("Microsoft YaHei", 10, "bold")
).pack(side=tk.LEFT, padx=3)

tk.Button(
    btn_traj_input,
    text="读取当前TCP并写入",
    command=read_current_tcp_to_traj,
    width=20
).pack(side=tk.LEFT, padx=3)

tk.Button(
    btn_traj_input,
    text="读取当前关节并写入",
    command=read_current_joints_to_traj,
    width=20
).pack(side=tk.LEFT, padx=3)

tk.Button(
    btn_traj_input,
    text="清空当前输入",
    command=clear_trajectory_input,
    width=16
).pack(side=tk.LEFT, padx=3)

tk.Label(
    tab_traj,
    text="加入点时检查格式并保留关节圈数；执行前再进行整段限位、台子和地面碰撞检查。",
    fg="#555555"
).pack(anchor=tk.W, padx=15, pady=3)

frame_record = tk.LabelFrame(
    tab_traj,
    text="已检查通过的连续运动点（按加入顺序执行，可混合 TCP / 关节点）"
)
frame_record.pack(fill=tk.BOTH, expand=True, padx=10, pady=8)

record_text = tk.Text(frame_record, font=("Consolas", 10), height=10)
record_text.pack(fill=tk.BOTH, expand=True, padx=5, pady=5)

btn_record_frame = tk.Frame(tab_traj)
btn_record_frame.pack(fill=tk.X, padx=10, pady=4)

tk.Button(
    btn_record_frame, text="删除最后一点",
    command=delete_last_record, width=15
).pack(side=tk.LEFT, padx=3)

tk.Button(
    btn_record_frame, text="清空全部点",
    command=clear_records, width=15
).pack(side=tk.LEFT, padx=3)

tk.Button(
    btn_record_frame, text="导入轨迹",
    command=import_trajectory, width=14
).pack(side=tk.LEFT, padx=3)

tk.Button(
    btn_record_frame, text="执行整段连续运动",
    command=execute_recorded_trajectory,
    width=24,
    font=("Microsoft YaHei", 10, "bold"),
    bg="#4CAF50", fg="white"
).pack(side=tk.LEFT, padx=3)

tk.Label(
    tab_traj,
    text="执行前按实机当前关节完成台子/地面预检；仅执行已验证方案。驱动报断连时复核实际到位；未到位或其他异常时中止。",
    fg="#555555"
).pack(anchor=tk.W, padx=15, pady=4)

real_deviation_var = tk.StringVar(value="500.0")
frame_deviation = tk.Frame(root)
frame_deviation.pack(fill=tk.X, padx=10, pady=3)
tk.Label(frame_deviation, text="预检MoveJ兜底最大TCP偏离(mm)：").pack(side=tk.LEFT)
tk.Entry(frame_deviation, textvariable=real_deviation_var, width=10).pack(side=tk.LEFT)
tk.Label(frame_deviation, text="默认500：与TCP仿真/轨迹7~11验证口径一致；实机速度10 mm/s（v14w25 调慢）").pack(side=tk.LEFT, padx=8)

# v14w24：法兰补偿MOVL 默认开启，勾选框移除（工艺定型）。v14l 实机判决驱动 MOVL 无工具
# 补偿（按法兰执行，无补偿直发已拉黑勿回归）；v14p 将错就错把法兰位姿当笛卡尔目标直发，
# 法兰被精确送达→物理尖端走在认证直线上。v14w36/37：位姿由调用方自算 invH(PoseFrame)*SolveFK
# （动画=认证直线，根治关节弧假碰撞冻死），发送窗口配单位变换（校验/数字=法兰空间）。
# 适用：MoveL 细分段≤210mm 且姿态恒定（v14w35 门禁）；规划/预检/几何零改动；失败指纹照旧即停；净化失败自动回落细分。
real_movldirect_var = tk.BooleanVar(value=True)   # 仅保留变量接口（执行入口读取）；无 GUI 控件

# ---- 日志区 ----
frame_log = tk.LabelFrame(root, text="日志")
frame_log.pack(fill=tk.BOTH, expand=True, padx=10, pady=5)

text_log = scrolledtext.ScrolledText(frame_log, font=("Consolas", 10), height=8)
text_log.pack(fill=tk.BOTH, expand=True, padx=5, pady=5)

# ============================================================
# 启动
# ============================================================
log("机器人: " + robot.Name())
log("程序就绪。" + LOG_VERSION + " ｜ 模式：RUNMODE_RUN_ROBOT + robot.Connect() ｜ 文件日志：" + LOG_PATH)
_ensure_canonical_tool()   # v14w17：启动守护（覆盖"加载了带归零工具的存档"场景）
log("单点：输入坐标 -> 检测可达性 -> 执行 MoveL/MoveJ")
log("目标关节：输入 J1~J6 -> 实机 MoveJ（不经过 TCP/Fanuc 转换和 IK）")
log("连续运动（P2P v14w41）：短直线段(≤210mm/姿态恒定)强制 MoveL 直走（工艺贴面平移不走 MoveJ 弧）；前视选解（换向可行性）+前视绑定执行；同位姿停顿不重选；弧碰退回 MoveL；死路分支救援+避障选解；换向碰撞自动换向（反方向坐标修复）/回绕/切分支/MoveL到场；首点种子枚举+整段重试；长运动不分瓣一指令直达（MoveL 仍细分，步长20mm；断连等待与重连并行——v14o 静默重连；v14w27 工具=182mm、v14w28 把手网格工作点=182、v14w29 圆柱挡板后移82、v14w30 直发到位阈5°、v14w32 J6±360换同角表示、v14w33 换姿段MoveJ直达、v14w34 换姿段判据修真位置差、v14w35 直发段长门禁210、v14w39 窗口全程+模型钉终点、v14w40 工具126+场景退26、v14w26 实机速度10mm/s、J4×J5自干涉组合区禁选(-40006)；法兰补偿MOVL 默认开（无勾选框）：短直线≤210mm 一指令直发+法兰级验收+MoveJ纠偏，净化失败自动回落细分）。")

def _log_pump():
    try:
        while True:
            text_log.insert(tk.END, _log_queue.get_nowait() + NL)
            text_log.see(tk.END)
    except Exception:
        pass
    root.after(100, _log_pump)


_close_requested = False


def _idle_tool_guard():
    if not _real_running and not _tool_window_depth:
        try:
            if _same_tool_pose(robot.PoseTool(), eye(4)):
                _ensure_canonical_tool()
            if _close_requested:
                root.destroy()
                return
        except Exception as exc:
            _file_log('工具空闲守护失败：' + str(exc))
    root.after(1000, _idle_tool_guard)


def _on_close():
    global _close_requested
    if _real_running:
        _close_requested = True
        log('已请求关闭：等待当前任务结束并恢复 TCP 后关闭窗口，继续保留到位监控。')
        return
    _ensure_canonical_tool()
    root.destroy()


root.protocol('WM_DELETE_WINDOW', _on_close)
root.after(100, _log_pump)
root.after(1000, _idle_tool_guard)
_start_heartbeat()
try:
    root.mainloop()
except BaseException:
    import traceback
    _file_log('FATAL mainloop: ' + traceback.format_exc())
    raise

--- Python program TCP真实运动_P2P版_16稳定版_替换前_20261104_095940 ---
# -*- coding: utf-8 -*-
"""
RoboDK 实机运动控制（基于 robodk_movej_diag.py 的成功模式）
- 单点：TCP 输入 -> IK 检测 -> MoveL/MoveJ 执行
- 连续轨迹：与TCP仿真同款（姿态退让、J6特异点±180°/自转360°、避障规划+缓存）
2026-10-09：连续运动逻辑对齐 机械臂TCP仿真_副本.py；预检偏离默认 50→500（与验证口径一致）
模式：RUNMODE_RUN_ROBOT + robot.Connect()
"""

from robodk.robolink import *
from robodk.robomath import *
import tkinter as tk
from tkinter import ttk, scrolledtext, filedialog
import time
import math
import json
import itertools

ROBOT_SPEED = 10.0   # v14w25：20→10 mm/s（用户要求调慢；顺带拉长指令间隔，缓解驱动掉线-重连压力）
CANONICAL_TOOL = (0.0, 0.0, 130.0, 0.0, 0.0, 0.0)   # v14w40：规范工具 182→126（2026-10-23 最终实测 法兰→TCP=126；v14w27~39 为 182、v14w14~w26 为 100）；守护用
NL = chr(10)
import queue as _queue_mod
_log_queue = _queue_mod.Queue()  # 后台线程日志经队列回流主线程，GUI 不冻结
LOG_PATH = r'D:\mydata\glm-workplace\sim_scripts\real_gui_log_p2p.txt'  # P2P版独立日志，不覆盖v13黑匣子
LOG_VERSION = 'v15.21-20261103'   # ★ 版本号规则（用户 2026-11-03 要求）：【每次改动都要升版本号】
                               # v15   ：从 v14w42 更名（J4 150→178 / P9 入禁直发 / Tool-User 实验开关 / 删超长横幅）
                               # v15.1 ：最后防线同角归一化修复（段6 J4=198.78 ≡ −161.22 被误判超限）
                               # v15.2 ：新增 |J4|>150 单独硬禁区（治 P5 的 J4=172.88 姿态自干涉）
                               # v15.3 ：打开 MOVL_SEND_TOOL_USER（直发前发 Tool(0)/User(0)，验证能否根治断断续续）
                               # v15.4 ：收口 MoveJ 加重试（治 P8 停下：收口遇断连没走完 ⇒ 关节残差 2.68° 残留）
                               # v15.5 ：直发+收口后再做【关节校正重试】（治 P8 停下：收口走假断连分支 ⇒ 报"已完成"但关节没到位）
                               # v15.6 ：_require_joints 改【带重试的稳定判定】（治 P8 尾通过 → P9 开头又失败：中间还在微动）
                               # v15.7 ：直发后先等【关节真静止】再做验收/收口（治 P8 的 elbow-flip 假通过/假失败）
                               # v15.8 ：★直发落点【自干涉安全网】—— 控制器自行选解可能落进禁区 ⇒ 立刻回认证构型
                               # v15.9 ：P8 也禁直发（治"选解自由"：J1/J6 同步偏 9.77° = 另一组 IK 解）⇒ P8 走细分
                               # v15.10：_require_joints 失败时【主动发 MoveJ 校正】（根治 P8 后不动：断连分支对 MoveJ 只等静止不等到位）
                               # 下次改动 ⇒ v15.22；标题与下方"连续运动"横幅要同步改
# v14w41：独立命名 TCP/法兰工具；恢复原工具链接并核验，失败停止；空闲守护与延后关闭。
# 历史版本记录（场景坐标并非实时状态）：★ v14w40（2026-10-23 18:09）：工具定案 126——最终实测 法兰→TCP=126，CANONICAL_TOOL/守护恢复值/banner 同步 126（历史：v14w27~39=182、v14w14~26=100）；配套场景 磨砂圆柱 y −860→−886、挡板 y 56→30（整体 −26 抵消工具加长的 26mm 深度偏移），轨迹13 采用 z460 统一版（连续轨迹13_t126_z460.json）——tool126+z460+场景−26 组合实测预检 21/21 PASS。⚠️ 实物圆柱/挡板须同步 −26；面贴滚轮旧坐标全部失效需重解；轨迹14/15 需在新配置下复验。v14w39（2026-10-22 14:31）：flange 窗口（单位变换+藏把手）从「仅包 RPC」扩大到【覆盖整个 settle 生命周期】。v14w38 失败教训：假断连让 MoveL 调用秒抛、窗口当场关闭、把手提前恢复，而真实滑行+RoboDK 本地退化动画仍在跑——本地动画在弧 66% 被碰撞检测掐停（模型冻点 J1≈67 四次实录同一位置）、红显常驻，收口 MoveJ 从撞点姿态发出被 RoboDK 拦死。v14w39 三件套：①窗口=包装层全程（发送+断连恢复+到位等待，补发重试每次重开窗）；②守卫补恢复隐藏态门把手（防 GUI 中杀留下隐藏态污染预检）；③直发 settle 返回后 robot.setJoints 钉模型到认证终点（清残余态双保险）。真直线 1mm 检查 0 碰撞、柜子零报警不变。v14w38：窗口藏把手（范围不足判负）。v14w37：位姿传递+单位变换（P8 TargetReachError 修复）。v14w35：门禁 210。v14w34：_seg_mm_ro 真位置差。其余见前版注释与 MEMORY。
# v14w32（2026-10-21 10:58）：J6 贴 ±360 边界的处置从「±359.999 内推」改为「换 (−180,180] 同角表示」（359.999→−0.001）——10-21 P4 实证：内推值仍被控制器丢 J6 单轴（J1~J5 全到、J6 停在 180、误差 180°）；换表示后当场重检 MoveJ 路径（方向翻转风险）；spin360/|J6|>360.001 不处理。其余=v14w30（阈值5°；v14w31 已撤回）。
# v14w30（2026-10-21 09:31）：MovL 直发到位阈 MOVL_ARRIVE_TOL_DEG 2°→5°——10-21 P8 实证：tool=182+z=380 构型下控制器 ~5mm 固有落点误差映射为关节 2.58°（tool=100 时代仅 0.7~0.9°），卡死在旧 ≤2° 阈值外被误判"疑似未执行"；臂实为完成态（零速/模式5/无报警）。护栏不降级：法兰级粗验收(≤8mm/≤1°)+MoveJ 收口仍在其后罩终点；60s 上限与不重发不变。（v14w31 稳定窗+补发×3 已于 10-21 按用户要求撤回。）
# v14w29（2026-10-20 16:42）：站内 圆柱+挡板 统一后移（远离基座）82mm（用户指令：尖端距圆柱面仅 14mm 太近、易自干涉）——圆柱 pose.y −840→−922、挡板 pose.y 76→−6；同时修正 10-15 起过期的场景注释。轨迹13 六点 z−82 补丁后离线预检 21/21 全绿（含本次场景移动复验）。
# v14w28（2026-10-20 16:15）：网格注释同步（纯注释版，逻辑零改动）——把手网格手术 v4：连接件加长、把手组件整体外移，【把手工作点=法兰前 182mm】，stl=tools\handle_rod_182_v2.stl（站内已换、未保存）。工具仍=182mm。
# v14w27（2026-10-20 15:49）：工具坐标 100→182mm（用户实测【物理工具真实长度】；站内 PoseTool 已同步 [0,0,182]）——CANONICAL_TOOL/守护恢复值/直发注释同步，全部 IK 按 182 解算。⚠️ 轨迹13 有 5 点（P8/P9/P10/P12/P13）在 182 下超臂展无逆解，重新示教前禁实机。
# v14w26（2026-10-15 18:15）：实机自干涉组合区（PoseSelfInterference 的 J4×J5 耦合，-40006 实录）——J4=-115.5×J5=173.1 与 J4=-109.4×J5=171.5 双拒；安全实录 J4=-83.2×J5=177.6。修：规划期禁选 |J4|>100 且 |J5|>165 的组合（MoveJ 解落区自动换无碰安全分支；直线段落区回落；无安全分支则整段换种子）。沿用 v14w25：速度10mm/s、J6±360内推（保留作防御）；v14w24：短直线强制MoveL、直发默认开。
# v14w20：受控补发。v14w19：三角离零域。v14w17：工具守护。工具=182.000（v14w27 起）；把手网格=v4 手术（把手组件外移、工作点 z=182，尖端=TCP，把手端抓手 z∈[174,182]；v14w28 起 stl=handle_rod_182_v2）。
# 场景（2026-10-20 实测，v14w29 圆柱/挡板统一后移82 后）：圆柱（轴∥X 滚轮 R150×H50）世界包络 X[−25,25] Y[−1062,−782] Z[330,610]；挡板世界包络 X[−235,215] Y[−1232,−932] Z[150,900]。10-13 版旧场景注释坐标已废（10-15 起站内多次平移未同步注释，v14w29 起以本行为准）。
# 控制器日志实锤（logs/all/log）：
#   11:38:20 拒收 MovL(-0.000000,-615.371000,300.000000,90.000000,0.000000,-0.000000)
#            → [MovL#820] the type of params is wrong: -30001 —— 这才是 P9 直发 60s 零位移的真凶；
#   15:55:51 单步同目标接受 MovL(0.000000,-615.371000,299.999986,89.999995,-0.000003,0.000000)
#            → return 0，1.1s 到位、法兰验收 5.08mm/0.61° 过。两样本差在【边界形态】：
#            x 负零/极小负、rx 恰=+90.000000、rz 负零（触发器三候选未最终定死，净化同时设防）。
# 修法：直发前 _movl_digit_safe_joints 只在零附近边界区对发送关节微扰（单关节 ≤0.05°、末端 ≲0.6mm
#   ≪ 圆柱真裕度 19.9mm）；到位/法兰验收/MoveJ 收口仍全部对【原始认证关节】判定，收口回认证构型。
#   净化失败 ⇒ 本段自动改走细分途经点（安全回落，不比 v14u 更糟）。
# 备份：…_v14v4_20261013-1608.py.bak（另有 1208 站内导出副本）；v14v/v2/v3 回退项见 P2P_LESSONS.md。
# 旧 v14u 备注：v14t 10:38 复跑判读——P9 起步延迟 >6s，「起点静止」与「完成静止」反馈不可区分，位置对目标才是唯一可靠锚点
# v12 黑匣子：原生崩溃时把 Python 调用栈转储到独立文件（被动，不影响逻辑）
# 注意：faulthandler.enable 只接受文件对象，传路径字符串会 AttributeError（v12 首版踩坑，已被 except 吞掉）
CRASH_PATH = r'D:\mydata\glm-workplace\sim_scripts\real_gui_crash.txt'
try:
    import faulthandler as _fh
    _crash_fp = open(CRASH_PATH, 'a', encoding='utf-8')
    _fh.enable(_crash_fp, all_threads=True)
except Exception:
    pass

def _file_log(s):
    try:
        import io as _io, time as _time
        with _io.open(LOG_PATH, 'a', encoding='utf-8') as f:
            f.write(_time.strftime('%m-%d %H:%M:%S') + ' | ' + str(s) + NL)
    except Exception:
        pass


RDK = Robolink()

def fanuc_to_pose(x, y, z, rx, ry, rz):
    return Fanuc_2_Pose([x, y, z, rx, ry, rz])

def pose_to_fanuc(pose):
    return Pose_2_Fanuc(pose)

# ---- 获取机器人 ----
robot = RDK.Item('Dobot CR5', ITEM_TYPE_ROBOT)
if not robot.Valid():
    raise Exception("未找到机器人")

# ---- 全局变量 ----
text_points = None
text_log = None
record_text = None
entries_single = None
entries_joint = None
move_type = None
trajectory_records = []
_connected = False

# ============================================================
# 日志
# ============================================================
# v12 心跳：每5秒覆写一次小文件（时间戳+pid+日志末行），进程死亡时间一目了然
HEARTBEAT_PATH = r'D:\mydata\glm-workplace\sim_scripts\real_gui_heartbeat.txt'

